(* IEC 61131-3 sources: plc-st-coding-agent/progress/evidence/f14_v14_remaining_20261113/jobs/codex_minimax-m27 (part 3) *)

(* ---- public-hard-05.patch_base_03.st ---- *)
(* ENGINEERING_CONTRACT *)
(*
  PUB001: Manual mode - button activates output while held, stop at limit switch or release.
          Manual outputs: retention=hold_until_button_release OR limit, reset=button_release OR limit_reached.
  PUB002: Emergency stop - all outputs OFF, all state cleared. No retention. Reset=EmergencyStop=TRUE.
  PUB003-PUB012: Single step mode - 8-step sequence, Start to advance each step.
          Step outputs: retention=hold_until_limit, reset=limit_reached OR mode_exit.
          Step index 1..8 maps to: Down→Grip→Up→Right→Down→Release→Up→Left→(repeat).
  PUB013-PUB014: Single cycle mode - auto-execute 8 steps on Start, stop at home.
          Same output retention as PUB003-PUB012. Cycle reset=mode_exit only.
  PUB015-PUB016: Continuous mode - same as single cycle but repeat after home.
          Cycle restart trigger: timer PT after home, if Start still asserted.
  PUB017: GripLimitSwitch/ReleaseLimitSwitch signal action completion (not position).
          Grip/Release output: activation=entry_unless_limit, retention=limit FALSE,
          deactivation=limit TRUE (same scan). No explicit reset input.
  PUB018: Caller guarantees mutually exclusive mode inputs.
  PUB019: Opposite-direction pairs (Up/Down, Left/Right) must never energize together.
          Implementation: output TRUE only when opposite limit is FALSE.
  PUB020: Single step confirmation = Start button release, not level.
*)
(* CONTRACT_RULES [] *)

TYPE ArmStep : INT (Idle := 0, Step1 := 1, Step2 := 2, Step3 := 3, Step4 := 4,
                     Step5 := 5, Step6 := 6, Step7 := 7, Step8 := 8)
END_TYPE;

FUNCTION_BLOCK ArmController
VAR_INPUT
    ManualMode       : BOOL;
    SingleStepMode   : BOOL;
    SingleCycleMode  : BOOL;
    ContinuousMode   : BOOL;
    EmergencyStop    : BOOL;
    Start            : BOOL;
    DownButton       : BOOL;
    UpButton         : BOOL;
    LeftButton       : BOOL;
    RightButton      : BOOL;
    GripButton       : BOOL;
    ReleaseButton    : BOOL;
    DownLimitSwitch  : BOOL;
    UpLimitSwitch    : BOOL;
    LeftLimitSwitch  : BOOL;
    RightLimitSwitch : BOOL;
    GripLimitSwitch  : BOOL;
    ReleaseLimitSwitch : BOOL;
END_VAR
VAR_OUTPUT
    MoveDown       : BOOL;
    MoveUp         : BOOL;
    MoveLeft       : BOOL;
    MoveRight      : BOOL;
    ActivateGrip   : BOOL;
    ActivateRelease : BOOL;
END_VAR
VAR
    tmp_CurrentStep   : ArmStep := ArmStep.Idle;
    tmp_StartTrigger  : BOOL;
    tmp_StartReleased : BOOL;
    tmp_Gripping      : BOOL;
    tmp_Releasing     : BOOL;
    tmp_CycleDoneTimer : TON;
END_VAR

// Emergency stop: clears all outputs and state
IF EmergencyStop THEN
    MoveDown       := FALSE;
    MoveUp         := FALSE;
    MoveLeft       := FALSE;
    MoveRight      := FALSE;
    ActivateGrip   := FALSE;
    ActivateRelease := FALSE;
    tmp_CurrentStep   := ArmStep.Idle;
    tmp_StartTrigger  := FALSE;
    tmp_StartReleased := FALSE;
    tmp_Gripping      := FALSE;
    tmp_Releasing     := FALSE;
    tmp_CycleDoneTimer(IN := FALSE, PT := T#0s);
    RETURN;
END_IF;

// Default all outputs OFF
MoveDown       := FALSE;
MoveUp         := FALSE;
MoveLeft       := FALSE;
MoveRight      := FALSE;
ActivateGrip   := FALSE;
ActivateRelease := FALSE;

IF ManualMode THEN
    // Direct button-to-output mapping, stop at limit switch
    MoveDown       := DownButton AND NOT DownLimitSwitch;
    MoveUp         := UpButton AND NOT UpLimitSwitch;
    MoveLeft       := LeftButton AND NOT LeftLimitSwitch;
    MoveRight      := RightButton AND NOT RightLimitSwitch;
    ActivateGrip   := GripButton AND NOT GripLimitSwitch;
    ActivateRelease := ReleaseButton AND NOT ReleaseLimitSwitch;

ELSIF SingleStepMode THEN
    // Rising-edge Start advances through steps; each step waits for limit switch
    IF tmp_StartReleased AND NOT Start AND tmp_CurrentStep = ArmStep.Idle THEN
        tmp_StartTrigger := TRUE;
    END_IF;
    tmp_StartReleased := Start;

    IF tmp_CurrentStep = ArmStep.Idle THEN
        IF tmp_StartTrigger THEN
            tmp_CurrentStep := ArmStep.Step1;
            tmp_StartTrigger := FALSE;
        END_IF;
    ELSE
        CASE TO_INT(tmp_CurrentStep) OF
            1: MoveDown := NOT DownLimitSwitch;
               IF DownLimitSwitch THEN
                   tmp_CurrentStep := ArmStep.Step2;
               END_IF;
            2: ActivateGrip := NOT GripLimitSwitch;
               IF GripLimitSwitch THEN
                   tmp_CurrentStep := ArmStep.Step3;
               END_IF;
            3: MoveUp := NOT UpLimitSwitch;
               IF UpLimitSwitch THEN
                   tmp_CurrentStep := ArmStep.Step4;
               END_IF;
            4: MoveRight := NOT RightLimitSwitch;
               IF RightLimitSwitch THEN
                   tmp_CurrentStep := ArmStep.Step5;
               END_IF;
            5: MoveDown := NOT DownLimitSwitch;
               IF DownLimitSwitch THEN
                   tmp_CurrentStep := ArmStep.Step6;
               END_IF;
            6: ActivateRelease := NOT ReleaseLimitSwitch;
               IF ReleaseLimitSwitch THEN
                   tmp_CurrentStep := ArmStep.Step7;
               END_IF;
            7: MoveUp := NOT UpLimitSwitch;
               IF UpLimitSwitch THEN
                   tmp_CurrentStep := ArmStep.Step8;
               END_IF;
            8: MoveLeft := NOT LeftLimitSwitch;
               IF LeftLimitSwitch THEN
                   tmp_CurrentStep := ArmStep.Idle;
               END_IF;
        END_CASE;
    END_IF;

ELSIF SingleCycleMode THEN
    // Start triggers auto-sequence; cycle completes and stops at home
    IF Start AND tmp_CurrentStep = ArmStep.Idle AND NOT tmp_Gripping AND NOT tmp_Releasing THEN
        tmp_StartTrigger := TRUE;
    END_IF;

    // Cycle completion: at Step8 and home (UpLimitSwitch AND LeftLimitSwitch)
    IF tmp_CurrentStep = ArmStep.Step8 AND UpLimitSwitch AND LeftLimitSwitch THEN
        tmp_CycleDoneTimer(IN := TRUE, PT := T#1ms);
        IF tmp_CycleDoneTimer.Q THEN
            tmp_StartTrigger  := FALSE;
            tmp_Gripping      := FALSE;
            tmp_Releasing     := FALSE;
            tmp_CurrentStep   := ArmStep.Idle;
        END_IF;
    ELSE
        tmp_CycleDoneTimer(IN := FALSE, PT := T#0s);
    END_IF;

    IF tmp_StartTrigger THEN
        CASE TO_INT(tmp_CurrentStep) OF
            0: tmp_CurrentStep := ArmStep.Step1;
            1: MoveDown := NOT DownLimitSwitch;
               IF DownLimitSwitch THEN
                   tmp_CurrentStep := ArmStep.Step2;
               END_IF;
            2: ActivateGrip := NOT GripLimitSwitch;
               IF GripLimitSwitch THEN
                   tmp_CurrentStep := ArmStep.Step3;
               END_IF;
            3: MoveUp := NOT UpLimitSwitch;
               IF UpLimitSwitch THEN
                   tmp_CurrentStep := ArmStep.Step4;
               END_IF;
            4: MoveRight := NOT RightLimitSwitch;
               IF RightLimitSwitch THEN
                   tmp_CurrentStep := ArmStep.Step5;
               END_IF;
            5: MoveDown := NOT DownLimitSwitch;
               IF DownLimitSwitch THEN
                   tmp_CurrentStep := ArmStep.Step6;
               END_IF;
            6: ActivateRelease := NOT ReleaseLimitSwitch;
               IF ReleaseLimitSwitch THEN
                   tmp_CurrentStep := ArmStep.Step7;
               END_IF;
            7: MoveUp := NOT UpLimitSwitch;
               IF UpLimitSwitch THEN
                   tmp_CurrentStep := ArmStep.Step8;
               END_IF;
            8: MoveLeft := NOT LeftLimitSwitch;
               IF LeftLimitSwitch THEN
                   tmp_CurrentStep := ArmStep.Idle;
               END_IF;
        END_CASE;
    END_IF;

ELSIF ContinuousMode THEN
    // Same as single cycle but restarts automatically after PT delay at home
    IF Start AND NOT tmp_Gripping AND NOT tmp_Releasing THEN
        tmp_StartTrigger := TRUE;
    END_IF;

    IF tmp_CurrentStep = ArmStep.Step8 AND UpLimitSwitch AND LeftLimitSwitch THEN
        tmp_CycleDoneTimer(IN := tmp_CycleDoneTimer.Q, PT := T#1ms);
        IF tmp_CycleDoneTimer.Q THEN
            tmp_CurrentStep := ArmStep.Idle;
        END_IF;
        IF NOT tmp_CycleDoneTimer.Q AND tmp_CurrentStep = ArmStep.Idle THEN
            tmp_StartTrigger := Start;
            tmp_Gripping     := FALSE;
            tmp_Releasing    := FALSE;
        END_IF;
    ELSE
        tmp_CycleDoneTimer(IN := FALSE, PT := T#0s);
    END_IF;

    IF tmp_StartTrigger THEN
        CASE TO_INT(tmp_CurrentStep) OF
            0: tmp_CurrentStep := ArmStep.Step1;
            1: MoveDown := NOT DownLimitSwitch;
               IF DownLimitSwitch THEN
                   tmp_CurrentStep := ArmStep.Step2;
               END_IF;
            2: ActivateGrip := NOT GripLimitSwitch;
               IF GripLimitSwitch THEN
                   tmp_CurrentStep := ArmStep.Step3;
               END_IF;
            3: MoveUp := NOT UpLimitSwitch;
               IF UpLimitSwitch THEN
                   tmp_CurrentStep := ArmStep.Step4;
               END_IF;
            4: MoveRight := NOT RightLimitSwitch;
               IF RightLimitSwitch THEN
                   tmp_CurrentStep := ArmStep.Step5;
               END_IF;
            5: MoveDown := NOT DownLimitSwitch;
               IF DownLimitSwitch THEN
                   tmp_CurrentStep := ArmStep.Step6;
               END_IF;
            6: ActivateRelease := NOT ReleaseLimitSwitch;
               IF ReleaseLimitSwitch THEN
                   tmp_CurrentStep := ArmStep.Step7;
               END_IF;
            7: MoveUp := NOT UpLimitSwitch;
               IF UpLimitSwitch THEN
                   tmp_CurrentStep := ArmStep.Step8;
               END_IF;
            8: MoveLeft := NOT LeftLimitSwitch;
               IF LeftLimitSwitch THEN
                   tmp_CurrentStep := ArmStep.Idle;
               END_IF;
        END_CASE;
    END_IF;
END_IF;

END_FUNCTION_BLOCK

(* ---- public-hard-05.raw_candidate_01.st ---- *)
(* ENGINEERING_CONTRACT *)
(*
  PUB001: Manual mode - button activates output while held, stop at limit switch or release.
          Manual outputs: retention=hold_until_button_release OR limit, reset=button_release OR limit_reached.
  PUB002: Emergency stop - all outputs OFF, all state cleared. No retention. Reset=EmergencyStop=TRUE.
  PUB003-PUB012: Single step mode - 8-step sequence, Start to advance each step.
          Step outputs: retention=hold_until_limit, reset=limit_reached OR mode_exit.
          Step index 1..8 maps to: Down→Grip→Up→Right→Down→Release→Up→Left→(repeat).
  PUB013-PUB014: Single cycle mode - auto-execute 8 steps on Start, stop at home.
          Same output retention as PUB003-PUB012. Cycle reset=mode_exit only.
  PUB015-PUB016: Continuous mode - same as single cycle but repeat after home.
          Cycle restart trigger: timer PT after home, if Start still asserted.
  PUB017: GripLimitSwitch/ReleaseLimitSwitch signal action completion (not position).
          Grip/Release output: activation=entry_unless_limit, retention=limit FALSE,
          deactivation=limit TRUE (same scan). No explicit reset input.
  PUB018: Caller guarantees mutually exclusive mode inputs.
  PUB019: Opposite-direction pairs (Up/Down, Left/Right) must never energize together.
          Implementation: output TRUE only when opposite limit is FALSE.
  PUB020: Single step confirmation = Start button release, not level.
*)
(* CONTRACT_RULES [] *)

TYPE ArmStep : INT (Idle := 0, Step1 := 1, Step2 := 2, Step3 := 3, Step4 := 4,
                     Step5 := 5, Step6 := 6, Step7 := 7, Step8 := 8)
END_TYPE

FUNCTION_BLOCK ArmController
VAR_INPUT
    ManualMode       : BOOL;
    SingleStepMode   : BOOL;
    SingleCycleMode  : BOOL;
    ContinuousMode   : BOOL;
    EmergencyStop    : BOOL;
    Start            : BOOL;
    DownButton       : BOOL;
    UpButton         : BOOL;
    LeftButton       : BOOL;
    RightButton      : BOOL;
    GripButton       : BOOL;
    ReleaseButton    : BOOL;
    DownLimitSwitch  : BOOL;
    UpLimitSwitch    : BOOL;
    LeftLimitSwitch  : BOOL;
    RightLimitSwitch : BOOL;
    GripLimitSwitch  : BOOL;
    ReleaseLimitSwitch : BOOL;
END_VAR
VAR_OUTPUT
    MoveDown       : BOOL;
    MoveUp         : BOOL;
    MoveLeft       : BOOL;
    MoveRight      : BOOL;
    ActivateGrip   : BOOL;
    ActivateRelease : BOOL;
END_VAR
VAR
    tmp_CurrentStep   : ArmStep := ArmStep.Idle;
    tmp_StartTrigger  : BOOL;
    tmp_StartReleased : BOOL;
    tmp_Gripping      : BOOL;
    tmp_Releasing     : BOOL;
    tmp_CycleDoneTimer : TON;
END_VAR

// Emergency stop: clears all outputs and state
IF EmergencyStop THEN
    MoveDown       := FALSE;
    MoveUp         := FALSE;
    MoveLeft       := FALSE;
    MoveRight      := FALSE;
    ActivateGrip   := FALSE;
    ActivateRelease := FALSE;
    tmp_CurrentStep   := ArmStep.Idle;
    tmp_StartTrigger  := FALSE;
    tmp_StartReleased := FALSE;
    tmp_Gripping      := FALSE;
    tmp_Releasing     := FALSE;
    tmp_CycleDoneTimer(IN := FALSE, PT := T#0s);
    RETURN;
END_IF;

// Default all outputs OFF
MoveDown       := FALSE;
MoveUp         := FALSE;
MoveLeft       := FALSE;
MoveRight      := FALSE;
ActivateGrip   := FALSE;
ActivateRelease := FALSE;

IF ManualMode THEN
    // Direct button-to-output mapping, stop at limit switch
    MoveDown       := DownButton AND NOT DownLimitSwitch;
    MoveUp         := UpButton AND NOT UpLimitSwitch;
    MoveLeft       := LeftButton AND NOT LeftLimitSwitch;
    MoveRight      := RightButton AND NOT RightLimitSwitch;
    ActivateGrip   := GripButton AND NOT GripLimitSwitch;
    ActivateRelease := ReleaseButton AND NOT ReleaseLimitSwitch;

ELSIF SingleStepMode THEN
    // Rising-edge Start advances through steps; each step waits for limit switch
    IF tmp_StartReleased AND NOT Start AND tmp_CurrentStep = ArmStep.Idle THEN
        tmp_StartTrigger := TRUE;
    END_IF
    tmp_StartReleased := Start;

    IF tmp_CurrentStep = ArmStep.Idle THEN
        IF tmp_StartTrigger THEN
            tmp_CurrentStep := ArmStep.Step1;
            tmp_StartTrigger := FALSE;
        END_IF;
    ELSE
        CASE TO_INT(tmp_CurrentStep) OF
            1: MoveDown := NOT DownLimitSwitch;
               IF DownLimitSwitch THEN
                   tmp_CurrentStep := ArmStep.Step2;
               END_IF;
            2: ActivateGrip := NOT GripLimitSwitch;
               IF GripLimitSwitch THEN
                   tmp_CurrentStep := ArmStep.Step3;
               END_IF;
            3: MoveUp := NOT UpLimitSwitch;
               IF UpLimitSwitch THEN
                   tmp_CurrentStep := ArmStep.Step4;
               END_IF;
            4: MoveRight := NOT RightLimitSwitch;
               IF RightLimitSwitch THEN
                   tmp_CurrentStep := ArmStep.Step5;
               END_IF;
            5: MoveDown := NOT DownLimitSwitch;
               IF DownLimitSwitch THEN
                   tmp_CurrentStep := ArmStep.Step6;
               END_IF;
            6: ActivateRelease := NOT ReleaseLimitSwitch;
               IF ReleaseLimitSwitch THEN
                   tmp_CurrentStep := ArmStep.Step7;
               END_IF;
            7: MoveUp := NOT UpLimitSwitch;
               IF UpLimitSwitch THEN
                   tmp_CurrentStep := ArmStep.Step8;
               END_IF;
            8: MoveLeft := NOT LeftLimitSwitch;
               IF LeftLimitSwitch THEN
                   tmp_CurrentStep := ArmStep.Idle;
               END_IF;
        END_CASE;
    END_IF;

ELSIF SingleCycleMode THEN
    // Start triggers auto-sequence; cycle completes and stops at home
    IF Start AND tmp_CurrentStep = ArmStep.Idle AND NOT tmp_Gripping AND NOT tmp_Releasing THEN
        tmp_StartTrigger := TRUE;
    END_IF;

    // Cycle completion: at Step8 and home (UpLimitSwitch AND LeftLimitSwitch)
    IF tmp_CurrentStep = ArmStep.Step8 AND UpLimitSwitch AND LeftLimitSwitch THEN
        tmp_CycleDoneTimer(IN := TRUE, PT := T#1ms);
        IF tmp_CycleDoneTimer.Q THEN
            tmp_StartTrigger  := FALSE;
            tmp_Gripping      := FALSE;
            tmp_Releasing     := FALSE;
            tmp_CurrentStep   := ArmStep.Idle;
        END_IF;
    ELSE
        tmp_CycleDoneTimer(IN := FALSE, PT := T#0s);
    END_IF;

    IF tmp_StartTrigger THEN
        CASE TO_INT(tmp_CurrentStep) OF
            0: tmp_CurrentStep := ArmStep.Step1;
            1: MoveDown := NOT DownLimitSwitch;
               IF DownLimitSwitch THEN
                   tmp_CurrentStep := ArmStep.Step2;
               END_IF;
            2: ActivateGrip := NOT GripLimitSwitch;
               IF GripLimitSwitch THEN
                   tmp_CurrentStep := ArmStep.Step3;
               END_IF;
            3: MoveUp := NOT UpLimitSwitch;
               IF UpLimitSwitch THEN
                   tmp_CurrentStep := ArmStep.Step4;
               END_IF;
            4: MoveRight := NOT RightLimitSwitch;
               IF RightLimitSwitch THEN
                   tmp_CurrentStep := ArmStep.Step5;
               END_IF;
            5: MoveDown := NOT DownLimitSwitch;
               IF DownLimitSwitch THEN
                   tmp_CurrentStep := ArmStep.Step6;
               END_IF;
            6: ActivateRelease := NOT ReleaseLimitSwitch;
               IF ReleaseLimitSwitch THEN
                   tmp_CurrentStep := ArmStep.Step7;
               END_IF;
            7: MoveUp := NOT UpLimitSwitch;
               IF UpLimitSwitch THEN
                   tmp_CurrentStep := ArmStep.Step8;
               END_IF;
            8: MoveLeft := NOT LeftLimitSwitch;
               IF LeftLimitSwitch THEN
                   tmp_CurrentStep := ArmStep.Idle;
               END_IF;
        END_CASE;
    END_IF;

ELSIF ContinuousMode THEN
    // Same as single cycle but restarts automatically after PT delay at home
    IF Start AND NOT tmp_Gripping AND NOT tmp_Releasing THEN
        tmp_StartTrigger := TRUE;
    END_IF;

    IF tmp_CurrentStep = ArmStep.Step8 AND UpLimitSwitch AND LeftLimitSwitch THEN
        tmp_CycleDoneTimer(IN := tmp_CycleDoneTimer.Q, PT := T#1ms);
        IF tmp_CycleDoneTimer.Q THEN
            tmp_CurrentStep := ArmStep.Idle;
        END_IF;
        IF NOT tmp_CycleDoneTimer.Q AND tmp_CurrentStep = ArmStep.Idle THEN
            tmp_StartTrigger := Start;
            tmp_Gripping     := FALSE;
            tmp_Releasing    := FALSE;
        END_IF;
    ELSE
        tmp_CycleDoneTimer(IN := FALSE, PT := T#0s);
    END_IF;

    IF tmp_StartTrigger THEN
        CASE TO_INT(tmp_CurrentStep) OF
            0: tmp_CurrentStep := ArmStep.Step1;
            1: MoveDown := NOT DownLimitSwitch;
               IF DownLimitSwitch THEN
                   tmp_CurrentStep := ArmStep.Step2;
               END_IF;
            2: ActivateGrip := NOT GripLimitSwitch;
               IF GripLimitSwitch THEN
                   tmp_CurrentStep := ArmStep.Step3;
               END_IF;
            3: MoveUp := NOT UpLimitSwitch;
               IF UpLimitSwitch THEN
                   tmp_CurrentStep := ArmStep.Step4;
               END_IF;
            4: MoveRight := NOT RightLimitSwitch;
               IF RightLimitSwitch THEN
                   tmp_CurrentStep := ArmStep.Step5;
               END_IF;
            5: MoveDown := NOT DownLimitSwitch;
               IF DownLimitSwitch THEN
                   tmp_CurrentStep := ArmStep.Step6;
               END_IF;
            6: ActivateRelease := NOT ReleaseLimitSwitch;
               IF ReleaseLimitSwitch THEN
                   tmp_CurrentStep := ArmStep.Step7;
               END_IF;
            7: MoveUp := NOT UpLimitSwitch;
               IF UpLimitSwitch THEN
                   tmp_CurrentStep := ArmStep.Step8;
               END_IF;
            8: MoveLeft := NOT LeftLimitSwitch;
               IF LeftLimitSwitch THEN
                   tmp_CurrentStep := ArmStep.Idle;
               END_IF;
        END_CASE;
    END_IF;
END_IF;

END_FUNCTION_BLOCK

(* ---- public-hard-06.candidate_01.st ---- *)
(*
ENGINEERING_CONTRACT
===================
PUB001: Mode 0=Manual, 1=Automatic (VAR_INPUT Mode)
PUB003: Manual interlock - ForwardButton→MotorForward, ReverseButton→MotorReverse, mutually exclusive
PUB002: Automatic sequential transport: Feed→Wash→Weigh→Fire→Output stations
PUB004: Station arrival detected by sensors; motor stops, awaits completion signal, then advances
PUB006: Weight qualification: qualified if 100<=weight<=200; else kick initiated
PUB007: FiringTemp calculation: weight[100,200]→temp[500,550] via linear interpolation
PUB008: CompletionLight ON when product detected at output, OFF when product removed
PUB005/P UB009-PUB012: washComplete/weightComplete/firingComplete are external process signals

OUTPUT STATE RETENTION
- MotorForward/MotorReverse: combinational per Mode selection, no retention across modes
- kick: pulse on weight qualification failure, no hold required
- CompletionLight: retained based on SensorOutput (hold until product removed)
- firingTemp: retained value written at weight station, held through firing until output

SCAN BEHAVIOR
- Sequential automatic states evaluate same-scan final state before output
- TON not required; all timing handled externally via completion signals
- Direction rule: MotorForward and MotorReverse never energized together
*)

FUNCTION_BLOCK ProductionControl
VAR_INPUT
    Mode            : BOOL;
    ForwardButton   : BOOL;
    ReverseButton   : BOOL;
    SensorFeed      : BOOL;
    SensorWash      : BOOL;
    SensorWeight    : BOOL;
    SensorFiring    : BOOL;
    SensorOutput    : BOOL;
    washComplete    : BOOL;
    weightComplete  : BOOL;
    weight          : REAL;
    firingComplete  : BOOL;
END_VAR

VAR_OUTPUT
    MotorForward    : BOOL;
    MotorReverse    : BOOL;
    kick             : BOOL;
    CompletionLight  : BOOL;
    firingTemp       : REAL;
END_VAR

VAR
    stepPosition    : INT := 0;
    localKick       : BOOL := FALSE;
END_VAR

(* CONTRACT_RULES [] *)

CASE stepPosition OF
    0: (* At feed station - waiting for material *)
        IF SensorFeed THEN
            MotorForward := TRUE;
            stepPosition := 1;
        END_IF;

    1: (* Moving to wash station - detecting arrival *)
        IF SensorWash THEN
            MotorForward := FALSE;
            stepPosition := 2;
        END_IF;

    2: (* At wash station - waiting for washComplete *)
        IF washComplete THEN
            MotorForward := TRUE;
            stepPosition := 3;
        END_IF;

    3: (* Moving to weight station - detecting arrival *)
        IF SensorWeight THEN
            MotorForward := FALSE;
            stepPosition := 4;
        END_IF;

    4: (* At weight station - waiting for weightComplete *)
        IF weightComplete THEN
            IF (weight >= 100.0) AND (weight <= 200.0) THEN
                firingTemp := 500.0 + (weight - 100.0) * (50.0 / 100.0);
                MotorForward := TRUE;
                stepPosition := 5;
            ELSE
                localKick := TRUE;
                kick := TRUE;
                MotorReverse := TRUE;
                stepPosition := 6;
            END_IF;
        END_IF;

    5: (* Moving to firing station - detecting arrival *)
        IF SensorFiring THEN
            MotorForward := FALSE;
            stepPosition := 7;
        END_IF;

    6: (* Rejection - returning to feed station *)
        localKick := FALSE;
        kick := FALSE;
        IF NOT SensorFeed THEN
            MotorReverse := FALSE;
            stepPosition := 0;
        END_IF;

    7: (* At firing station - waiting for firingComplete *)
        IF firingComplete THEN
            MotorForward := TRUE;
            stepPosition := 8;
        END_IF;

    8: (* Moving to output station - detecting arrival *)
        IF SensorOutput THEN
            MotorForward := FALSE;
            stepPosition := 9;
        END_IF;

    9: (* At output station - waiting for product removal *)
        CompletionLight := TRUE;

    ELSE
        stepPosition := 0;
END_CASE;

IF Mode = 0 THEN
    stepPosition := 0;
    MotorForward := FALSE;
    MotorReverse := FALSE;
    kick := FALSE;
    CompletionLight := FALSE;
    localKick := FALSE;
    firingTemp := 0.0;

    IF ForwardButton AND NOT ReverseButton THEN
        MotorForward := TRUE;
    ELSIF ReverseButton AND NOT ForwardButton THEN
        MotorReverse := TRUE;
    END_IF;
END_IF;

IF NOT SensorOutput AND stepPosition = 9 THEN
    CompletionLight := FALSE;
    stepPosition := 0;
END_IF;

END_FUNCTION_BLOCK

(* ---- public-hard-06.raw_candidate_01.st ---- *)
(*
ENGINEERING_CONTRACT
===================
PUB001: Mode 0=Manual, 1=Automatic (VAR_INPUT Mode)
PUB003: Manual interlock - ForwardButton→MotorForward, ReverseButton→MotorReverse, mutually exclusive
PUB002: Automatic sequential transport: Feed→Wash→Weigh→Fire→Output stations
PUB004: Station arrival detected by sensors; motor stops, awaits completion signal, then advances
PUB006: Weight qualification: qualified if 100<=weight<=200; else kick initiated
PUB007: FiringTemp calculation: weight[100,200]→temp[500,550] via linear interpolation
PUB008: CompletionLight ON when product detected at output, OFF when product removed
PUB005/P UB009-PUB012: washComplete/weightComplete/firingComplete are external process signals

OUTPUT STATE RETENTION
- MotorForward/MotorReverse: combinational per Mode selection, no retention across modes
- kick: pulse on weight qualification failure, no hold required
- CompletionLight: retained based on SensorOutput (hold until product removed)
- firingTemp: retained value written at weight station, held through firing until output

SCAN BEHAVIOR
- Sequential automatic states evaluate same-scan final state before output
- TON not required; all timing handled externally via completion signals
- Direction rule: MotorForward and MotorReverse never energized together
*)

FUNCTION_BLOCK ProductionControl
VAR_INPUT
    Mode            : BOOL;
    ForwardButton   : BOOL;
    ReverseButton   : BOOL;
    SensorFeed      : BOOL;
    SensorWash      : BOOL;
    SensorWeight    : BOOL;
    SensorFiring    : BOOL;
    SensorOutput    : BOOL;
    washComplete    : BOOL;
    weightComplete  : BOOL;
    weight          : REAL;
    firingComplete  : BOOL;
END_VAR

VAR_OUTPUT
    MotorForward    : BOOL;
    MotorReverse    : BOOL;
    kick             : BOOL;
    CompletionLight  : BOOL;
    firingTemp       : REAL;
END_VAR

VAR
    stepPosition    : INT := 0;
    localKick       : BOOL := FALSE;
END_VAR

(* CONTRACT_RULES [] *)

CASE stepPosition OF
    0: (* At feed station - waiting for material *)
        IF SensorFeed THEN
            MotorForward := TRUE;
            stepPosition := 1;
        END_IF

    1: (* Moving to wash station - detecting arrival *)
        IF SensorWash THEN
            MotorForward := FALSE;
            stepPosition := 2;
        END_IF

    2: (* At wash station - waiting for washComplete *)
        IF washComplete THEN
            MotorForward := TRUE;
            stepPosition := 3;
        END_IF

    3: (* Moving to weight station - detecting arrival *)
        IF SensorWeight THEN
            MotorForward := FALSE;
            stepPosition := 4;
        END_IF

    4: (* At weight station - waiting for weightComplete *)
        IF weightComplete THEN
            IF (weight >= 100.0) AND (weight <= 200.0) THEN
                firingTemp := 500.0 + (weight - 100.0) * (50.0 / 100.0);
                MotorForward := TRUE;
                stepPosition := 5;
            ELSE
                localKick := TRUE;
                kick := TRUE;
                MotorReverse := TRUE;
                stepPosition := 6;
            END_IF
        END_IF

    5: (* Moving to firing station - detecting arrival *)
        IF SensorFiring THEN
            MotorForward := FALSE;
            stepPosition := 7;
        END_IF

    6: (* Rejection - returning to feed station *)
        localKick := FALSE;
        kick := FALSE;
        IF NOT SensorFeed THEN
            MotorReverse := FALSE;
            stepPosition := 0;
        END_IF

    7: (* At firing station - waiting for firingComplete *)
        IF firingComplete THEN
            MotorForward := TRUE;
            stepPosition := 8;
        END_IF

    8: (* Moving to output station - detecting arrival *)
        IF SensorOutput THEN
            MotorForward := FALSE;
            stepPosition := 9;
        END_IF

    9: (* At output station - waiting for product removal *)
        CompletionLight := TRUE;

    ELSE
        stepPosition := 0;
END_CASE

IF Mode = 0 THEN
    stepPosition := 0;
    MotorForward := FALSE;
    MotorReverse := FALSE;
    kick := FALSE;
    CompletionLight := FALSE;
    localKick := FALSE;
    firingTemp := 0.0;

    IF ForwardButton AND NOT ReverseButton THEN
        MotorForward := TRUE;
    ELSIF ReverseButton AND NOT ForwardButton THEN
        MotorReverse := TRUE;
    END_IF
END_IF

IF NOT SensorOutput AND stepPosition = 9 THEN
    CompletionLight := FALSE;
    stepPosition := 0;
END_IF

END_FUNCTION_BLOCK

(* ---- public-medium-01.candidate_01.st ---- *)
FUNCTION_BLOCK FB_MultiPumpControl
VAR_INPUT
    mode : BOOL;          // FALSE: Manual mode, TRUE: Automatic mode
    start : BOOL;         // Start button
    stop : BOOL;          // Stop button
END_VAR

VAR_IN_OUT
    pumpGroup : ARRAY[1..5] OF ST_Pump;
END_VAR

VAR
    startRisingEdge : BOOL;               // Rising edge of start
    tmp_startPrev : BOOL;                 // Previous start state
    tmp_i : INT;                          // Loop counter
    tmp_j : INT;                          // Loop counter
    tmp_swap : INT;                       // Swap variable
    tmp_pumpIdx : ARRAY[1..5] OF INT;    // Pump indices for sorting
    tmp_priorities : ARRAY[1..5] OF INT; // Priority copy for sorting
    tmp_swap_idx : INT;                   // Index swap
END_VAR

// ENGINEERING_CONTRACT:
// PUB001 [L91-265]: mode=FALSE → manual; start activates pumps where selection=TRUE
// PUB001 [L91-265]: mode=TRUE → automatic; start activates top-3 by priority (3-in-2-standby)
// PUB002 [L266-350]: stop halts all pumps; no retention on stop (level-triggered)
// PUB003 [L351-463]: Rising edge on start evaluates selection; stop has same-scan priority
// PUB004 [L464-652]: Only RunComd is written; priority/selection are read-only

(* CONTRACT_RULES [] *)

startRisingEdge := start AND NOT tmp_startPrev;

IF stop THEN
    FOR tmp_i := 1 TO 5 DO
        pumpGroup[tmp_i].RunComd := FALSE;
    END_FOR;
ELSIF startRisingEdge THEN
    IF mode = FALSE THEN
        FOR tmp_i := 1 TO 5 DO
            IF pumpGroup[tmp_i].selection THEN
                pumpGroup[tmp_i].RunComd := TRUE;
            END_IF;
        END_FOR;
    ELSE
        FOR tmp_i := 1 TO 5 DO
            tmp_priorities[tmp_i] := pumpGroup[tmp_i].priority;
            tmp_pumpIdx[tmp_i] := tmp_i;
        END_FOR;
        FOR tmp_i := 1 TO 4 DO
            FOR tmp_j := tmp_i + 1 TO 5 DO
                IF tmp_priorities[tmp_j] > tmp_priorities[tmp_i] THEN
                    tmp_swap := tmp_priorities[tmp_i];
                    tmp_priorities[tmp_i] := tmp_priorities[tmp_j];
                    tmp_priorities[tmp_j] := tmp_swap;
                    tmp_swap_idx := tmp_pumpIdx[tmp_i];
                    tmp_pumpIdx[tmp_i] := tmp_pumpIdx[tmp_j];
                    tmp_pumpIdx[tmp_j] := tmp_swap_idx;
                END_IF;
            END_FOR;
        END_FOR;
        FOR tmp_i := 1 TO 5 DO
            IF tmp_i <= 3 THEN
                pumpGroup[tmp_pumpIdx[tmp_i]].RunComd := TRUE;
            ELSE
                pumpGroup[tmp_pumpIdx[tmp_i]].RunComd := FALSE;
            END_IF;
        END_FOR;
    END_IF;
END_IF;

tmp_startPrev := start;
END_FUNCTION_BLOCK

(* ---- public-medium-01.candidate_03.st ---- *)
TYPE ST_Pump :
STRUCT
    priority : INT;
    selection : BOOL;
    RunComd : BOOL;
END_STRUCT
END_TYPE;

FUNCTION_BLOCK FB_MultiPumpControl
VAR_INPUT
    mode : BOOL;          // FALSE: Manual mode, TRUE: Automatic mode
    start : BOOL;         // Start button
    stop : BOOL;          // Stop button
END_VAR

VAR_IN_OUT
    pumpGroup : ARRAY[1..5] OF ST_Pump;
END_VAR

VAR
    startRisingEdge : BOOL;               // Rising edge of start
    tmp_startPrev : BOOL;                 // Previous start state
    tmp_i : INT;                          // Loop counter
    tmp_j : INT;                          // Loop counter
    tmp_swap : INT;                       // Swap variable
    tmp_pumpIdx : ARRAY[1..5] OF INT;    // Pump indices for sorting
    tmp_priorities : ARRAY[1..5] OF INT; // Priority copy for sorting
    tmp_swap_idx : INT;                   // Index swap
END_VAR

// ENGINEERING_CONTRACT:
// PUB001 [L91-265]: mode=FALSE → manual; start activates pumps where selection=TRUE
// PUB001 [L91-265]: mode=TRUE → automatic; start activates top-3 by priority (3-in-2-standby)
// PUB002 [L266-350]: stop halts all pumps; no retention on stop (level-triggered)
// PUB003 [L351-463]: Rising edge on start evaluates selection; stop has same-scan priority
// PUB004 [L464-652]: Only RunComd is written; priority/selection are read-only

(* CONTRACT_RULES [] *)

startRisingEdge := start AND NOT tmp_startPrev;

IF stop THEN
    FOR tmp_i := 1 TO 5 DO
        pumpGroup[tmp_i].RunComd := FALSE;
    END_FOR;
ELSIF startRisingEdge THEN
    IF mode = FALSE THEN
        FOR tmp_i := 1 TO 5 DO
            IF pumpGroup[tmp_i].selection THEN
                pumpGroup[tmp_i].RunComd := TRUE;
            END_IF;
        END_FOR;
    ELSE
        FOR tmp_i := 1 TO 5 DO
            tmp_priorities[tmp_i] := pumpGroup[tmp_i].priority;
            tmp_pumpIdx[tmp_i] := tmp_i;
        END_FOR;
        FOR tmp_i := 1 TO 4 DO
            FOR tmp_j := tmp_i + 1 TO 5 DO
                IF tmp_priorities[tmp_j] > tmp_priorities[tmp_i] THEN
                    tmp_swap := tmp_priorities[tmp_i];
                    tmp_priorities[tmp_i] := tmp_priorities[tmp_j];
                    tmp_priorities[tmp_j] := tmp_swap;
                    tmp_swap_idx := tmp_pumpIdx[tmp_i];
                    tmp_pumpIdx[tmp_i] := tmp_pumpIdx[tmp_j];
                    tmp_pumpIdx[tmp_j] := tmp_swap_idx;
                END_IF;
            END_FOR;
        END_FOR;
        FOR tmp_i := 1 TO 5 DO
            IF tmp_i <= 3 THEN
                pumpGroup[tmp_pumpIdx[tmp_i]].RunComd := TRUE;
            ELSE
                pumpGroup[tmp_pumpIdx[tmp_i]].RunComd := FALSE;
            END_IF;
        END_FOR;
    END_IF;
END_IF;

tmp_startPrev := start;
END_FUNCTION_BLOCK

(* ---- public-medium-01.patch_base_02.st ---- *)
FUNCTION_BLOCK FB_MultiPumpControl
VAR_INPUT
    mode : BOOL;          // FALSE: Manual mode, TRUE: Automatic mode
    start : BOOL;         // Start button
    stop : BOOL;          // Stop button
END_VAR

VAR_IN_OUT
    pumpGroup : ARRAY[1..5] OF ST_Pump;
END_VAR

VAR
    startRisingEdge : BOOL;               // Rising edge of start
    tmp_startPrev : BOOL;                 // Previous start state
    tmp_i : INT;                          // Loop counter
    tmp_j : INT;                          // Loop counter
    tmp_swap : INT;                       // Swap variable
    tmp_pumpIdx : ARRAY[1..5] OF INT;    // Pump indices for sorting
    tmp_priorities : ARRAY[1..5] OF INT; // Priority copy for sorting
    tmp_swap_idx : INT;                   // Index swap
END_VAR

// ENGINEERING_CONTRACT:
// PUB001 [L91-265]: mode=FALSE → manual; start activates pumps where selection=TRUE
// PUB001 [L91-265]: mode=TRUE → automatic; start activates top-3 by priority (3-in-2-standby)
// PUB002 [L266-350]: stop halts all pumps; no retention on stop (level-triggered)
// PUB003 [L351-463]: Rising edge on start evaluates selection; stop has same-scan priority
// PUB004 [L464-652]: Only RunComd is written; priority/selection are read-only

(* CONTRACT_RULES [] *)

startRisingEdge := start AND NOT tmp_startPrev;

IF stop THEN
    FOR tmp_i := 1 TO 5 DO
        pumpGroup[tmp_i].RunComd := FALSE;
    END_FOR;
ELSIF startRisingEdge THEN
    IF mode = FALSE THEN
        FOR tmp_i := 1 TO 5 DO
            IF pumpGroup[tmp_i].selection THEN
                pumpGroup[tmp_i].RunComd := TRUE;
            END_IF;
        END_FOR;
    ELSE
        FOR tmp_i := 1 TO 5 DO
            tmp_priorities[tmp_i] := pumpGroup[tmp_i].priority;
            tmp_pumpIdx[tmp_i] := tmp_i;
        END_FOR;
        FOR tmp_i := 1 TO 4 DO
            FOR tmp_j := tmp_i + 1 TO 5 DO
                IF tmp_priorities[tmp_j] > tmp_priorities[tmp_i] THEN
                    tmp_swap := tmp_priorities[tmp_i];
                    tmp_priorities[tmp_i] := tmp_priorities[tmp_j];
                    tmp_priorities[tmp_j] := tmp_swap;
                    tmp_swap_idx := tmp_pumpIdx[tmp_i];
                    tmp_pumpIdx[tmp_i] := tmp_pumpIdx[tmp_j];
                    tmp_pumpIdx[tmp_j] := tmp_swap_idx;
                END_IF;
            END_FOR;
        END_FOR;
        FOR tmp_i := 1 TO 5 DO
            IF tmp_i <= 3 THEN
                pumpGroup[tmp_pumpIdx[tmp_i]].RunComd := TRUE;
            ELSE
                pumpGroup[tmp_pumpIdx[tmp_i]].RunComd := FALSE;
            END_IF;
        END_FOR;
    END_IF;
END_IF;

tmp_startPrev := start;
END_FUNCTION_BLOCK

(* ---- public-medium-01.patch_base_03.st ---- *)
FUNCTION_BLOCK FB_MultiPumpControl
VAR_INPUT
    mode : BOOL;          // FALSE: Manual mode, TRUE: Automatic mode
    start : BOOL;         // Start button
    stop : BOOL;          // Stop button
END_VAR

VAR_IN_OUT
    pumpGroup : ARRAY[1..5] OF ST_Pump;
END_VAR

VAR
    startRisingEdge : BOOL;               // Rising edge of start
    tmp_startPrev : BOOL;                 // Previous start state
    tmp_i : INT;                          // Loop counter
    tmp_j : INT;                          // Loop counter
    tmp_swap : INT;                       // Swap variable
    tmp_pumpIdx : ARRAY[1..5] OF INT;    // Pump indices for sorting
    tmp_priorities : ARRAY[1..5] OF INT; // Priority copy for sorting
    tmp_swap_idx : INT;                   // Index swap
END_VAR

// ENGINEERING_CONTRACT:
// PUB001 [L91-265]: mode=FALSE → manual; start activates pumps where selection=TRUE
// PUB001 [L91-265]: mode=TRUE → automatic; start activates top-3 by priority (3-in-2-standby)
// PUB002 [L266-350]: stop halts all pumps; no retention on stop (level-triggered)
// PUB003 [L351-463]: Rising edge on start evaluates selection; stop has same-scan priority
// PUB004 [L464-652]: Only RunComd is written; priority/selection are read-only

(* CONTRACT_RULES [] *)

startRisingEdge := start AND NOT tmp_startPrev;

IF stop THEN
    FOR tmp_i := 1 TO 5 DO
        pumpGroup[tmp_i].RunComd := FALSE;
    END_FOR;
ELSIF startRisingEdge THEN
    IF mode = FALSE THEN
        FOR tmp_i := 1 TO 5 DO
            IF pumpGroup[tmp_i].selection THEN
                pumpGroup[tmp_i].RunComd := TRUE;
            END_IF;
        END_FOR;
    ELSE
        FOR tmp_i := 1 TO 5 DO
            tmp_priorities[tmp_i] := pumpGroup[tmp_i].priority;
            tmp_pumpIdx[tmp_i] := tmp_i;
        END_FOR;
        FOR tmp_i := 1 TO 4 DO
            FOR tmp_j := tmp_i + 1 TO 5 DO
                IF tmp_priorities[tmp_j] > tmp_priorities[tmp_i] THEN
                    tmp_swap := tmp_priorities[tmp_i];
                    tmp_priorities[tmp_i] := tmp_priorities[tmp_j];
                    tmp_priorities[tmp_j] := tmp_swap;
                    tmp_swap_idx := tmp_pumpIdx[tmp_i];
                    tmp_pumpIdx[tmp_i] := tmp_pumpIdx[tmp_j];
                    tmp_pumpIdx[tmp_j] := tmp_swap_idx;
                END_IF;
            END_FOR;
        END_FOR;
        FOR tmp_i := 1 TO 5 DO
            IF tmp_i <= 3 THEN
                pumpGroup[tmp_pumpIdx[tmp_i]].RunComd := TRUE;
            ELSE
                pumpGroup[tmp_pumpIdx[tmp_i]].RunComd := FALSE;
            END_IF;
        END_FOR;
    END_IF;
END_IF;

tmp_startPrev := start;
END_FUNCTION_BLOCK

(* ---- public-medium-01.patch_base_04.st ---- *)
TYPE ST_Pump :
STRUCT
    priority : INT;
    selection : BOOL;
    RunComd : BOOL;
END_STRUCT
END_TYPE;

FUNCTION_BLOCK FB_MultiPumpControl
VAR_INPUT
    mode : BOOL;          // FALSE: Manual mode, TRUE: Automatic mode
    start : BOOL;         // Start button
    stop : BOOL;          // Stop button
END_VAR

VAR_IN_OUT
    pumpGroup : ARRAY[1..5] OF ST_Pump;
END_VAR

VAR
    startRisingEdge : BOOL;               // Rising edge of start
    tmp_startPrev : BOOL;                 // Previous start state
    tmp_i : INT;                          // Loop counter
    tmp_j : INT;                          // Loop counter
    tmp_swap : INT;                       // Swap variable
    tmp_pumpIdx : ARRAY[1..5] OF INT;    // Pump indices for sorting
    tmp_priorities : ARRAY[1..5] OF INT; // Priority copy for sorting
    tmp_swap_idx : INT;                   // Index swap
END_VAR

// ENGINEERING_CONTRACT:
// PUB001 [L91-265]: mode=FALSE → manual; start activates pumps where selection=TRUE
// PUB001 [L91-265]: mode=TRUE → automatic; start activates top-3 by priority (3-in-2-standby)
// PUB002 [L266-350]: stop halts all pumps; no retention on stop (level-triggered)
// PUB003 [L351-463]: Rising edge on start evaluates selection; stop has same-scan priority
// PUB004 [L464-652]: Only RunComd is written; priority/selection are read-only

(* CONTRACT_RULES [] *)

startRisingEdge := start AND NOT tmp_startPrev;

IF stop THEN
    FOR tmp_i := 1 TO 5 DO
        pumpGroup[tmp_i].RunComd := FALSE;
    END_FOR;
ELSIF startRisingEdge THEN
    IF mode = FALSE THEN
        FOR tmp_i := 1 TO 5 DO
            IF pumpGroup[tmp_i].selection THEN
                pumpGroup[tmp_i].RunComd := TRUE;
            END_IF;
        END_FOR;
    ELSE
        FOR tmp_i := 1 TO 5 DO
            tmp_priorities[tmp_i] := pumpGroup[tmp_i].priority;
            tmp_pumpIdx[tmp_i] := tmp_i;
        END_FOR;
        FOR tmp_i := 1 TO 4 DO
            FOR tmp_j := tmp_i + 1 TO 5 DO
                IF tmp_priorities[tmp_j] > tmp_priorities[tmp_i] THEN
                    tmp_swap := tmp_priorities[tmp_i];
                    tmp_priorities[tmp_i] := tmp_priorities[tmp_j];
                    tmp_priorities[tmp_j] := tmp_swap;
                    tmp_swap_idx := tmp_pumpIdx[tmp_i];
                    tmp_pumpIdx[tmp_i] := tmp_pumpIdx[tmp_j];
                    tmp_pumpIdx[tmp_j] := tmp_swap_idx;
                END_IF;
            END_FOR;
        END_FOR;
        FOR tmp_i := 1 TO 5 DO
            IF tmp_i <= 3 THEN
                pumpGroup[tmp_pumpIdx[tmp_i]].RunComd := TRUE;
            ELSE
                pumpGroup[tmp_pumpIdx[tmp_i]].RunComd := FALSE;
            END_IF;
        END_FOR;
    END_IF;
END_IF;

tmp_startPrev := start;
END_FUNCTION_BLOCK

(* ---- public-medium-01.raw_candidate_01.st ---- *)
FUNCTION_BLOCK FB_MultiPumpControl
VAR_INPUT
    mode : BOOL;          // FALSE: Manual mode, TRUE: Automatic mode
    start : BOOL;         // Start button
    stop : BOOL;          // Stop button
END_VAR

VAR_IN_OUT
    pumpGroup : ARRAY[1..5] OF ST_Pump;
END_VAR

VAR
    startRisingEdge : BOOL;               // Rising edge of start
    tmp_startPrev : BOOL;                 // Previous start state
    tmp_i : INT;                          // Loop counter
    tmp_j : INT;                          // Loop counter
    tmp_swap : INT;                       // Swap variable
    tmp_pumpIdx : ARRAY[1..5] OF INT;    // Pump indices for sorting
    tmp_priorities : ARRAY[1..5] OF INT; // Priority copy for sorting
    tmp_swap_idx : INT;                   // Index swap
END_VAR

// ENGINEERING_CONTRACT:
// PUB001 [L91-265]: mode=FALSE → manual; start activates pumps where selection=TRUE
// PUB001 [L91-265]: mode=TRUE → automatic; start activates top-3 by priority (3-in-2-standby)
// PUB002 [L266-350]: stop halts all pumps; no retention on stop (level-triggered)
// PUB003 [L351-463]: Rising edge on start evaluates selection; stop has same-scan priority
// PUB004 [L464-652]: Only RunComd is written; priority/selection are read-only

(* CONTRACT_RULES [] *)

startRisingEdge := start AND NOT tmp_startPrev;

IF stop THEN
    FOR tmp_i := 1 TO 5 DO
        pumpGroup[tmp_i].RunComd := FALSE;
    END_FOR
ELSIF startRisingEdge THEN
    IF mode = FALSE THEN
        FOR tmp_i := 1 TO 5 DO
            IF pumpGroup[tmp_i].selection THEN
                pumpGroup[tmp_i].RunComd := TRUE;
            END_IF
        END_FOR
    ELSE
        FOR tmp_i := 1 TO 5 DO
            tmp_priorities[tmp_i] := pumpGroup[tmp_i].priority;
            tmp_pumpIdx[tmp_i] := tmp_i;
        END_FOR
        FOR tmp_i := 1 TO 4 DO
            FOR tmp_j := tmp_i + 1 TO 5 DO
                IF tmp_priorities[tmp_j] > tmp_priorities[tmp_i] THEN
                    tmp_swap := tmp_priorities[tmp_i];
                    tmp_priorities[tmp_i] := tmp_priorities[tmp_j];
                    tmp_priorities[tmp_j] := tmp_swap;
                    tmp_swap_idx := tmp_pumpIdx[tmp_i];
                    tmp_pumpIdx[tmp_i] := tmp_pumpIdx[tmp_j];
                    tmp_pumpIdx[tmp_j] := tmp_swap_idx;
                END_IF
            END_FOR
        END_FOR
        FOR tmp_i := 1 TO 5 DO
            IF tmp_i <= 3 THEN
                pumpGroup[tmp_pumpIdx[tmp_i]].RunComd := TRUE;
            ELSE
                pumpGroup[tmp_pumpIdx[tmp_i]].RunComd := FALSE;
            END_IF
        END_FOR
    END_IF
END_IF

tmp_startPrev := start;
END_FUNCTION_BLOCK

(* ---- public-medium-01.raw_candidate_03.st ---- *)
TYPE ST_Pump :
STRUCT
    priority : INT;
    selection : BOOL;
    RunComd : BOOL;
END_STRUCT
END_TYPE

FUNCTION_BLOCK FB_MultiPumpControl
VAR_INPUT
    mode : BOOL;          // FALSE: Manual mode, TRUE: Automatic mode
    start : BOOL;         // Start button
    stop : BOOL;          // Stop button
END_VAR

VAR_IN_OUT
    pumpGroup : ARRAY[1..5] OF ST_Pump;
END_VAR

VAR
    startRisingEdge : BOOL;               // Rising edge of start
    tmp_startPrev : BOOL;                 // Previous start state
    tmp_i : INT;                          // Loop counter
    tmp_j : INT;                          // Loop counter
    tmp_swap : INT;                       // Swap variable
    tmp_pumpIdx : ARRAY[1..5] OF INT;    // Pump indices for sorting
    tmp_priorities : ARRAY[1..5] OF INT; // Priority copy for sorting
    tmp_swap_idx : INT;                   // Index swap
END_VAR

// ENGINEERING_CONTRACT:
// PUB001 [L91-265]: mode=FALSE → manual; start activates pumps where selection=TRUE
// PUB001 [L91-265]: mode=TRUE → automatic; start activates top-3 by priority (3-in-2-standby)
// PUB002 [L266-350]: stop halts all pumps; no retention on stop (level-triggered)
// PUB003 [L351-463]: Rising edge on start evaluates selection; stop has same-scan priority
// PUB004 [L464-652]: Only RunComd is written; priority/selection are read-only

(* CONTRACT_RULES [] *)

startRisingEdge := start AND NOT tmp_startPrev;

IF stop THEN
    FOR tmp_i := 1 TO 5 DO
        pumpGroup[tmp_i].RunComd := FALSE;
    END_FOR;
ELSIF startRisingEdge THEN
    IF mode = FALSE THEN
        FOR tmp_i := 1 TO 5 DO
            IF pumpGroup[tmp_i].selection THEN
                pumpGroup[tmp_i].RunComd := TRUE;
            END_IF;
        END_FOR;
    ELSE
        FOR tmp_i := 1 TO 5 DO
            tmp_priorities[tmp_i] := pumpGroup[tmp_i].priority;
            tmp_pumpIdx[tmp_i] := tmp_i;
        END_FOR;
        FOR tmp_i := 1 TO 4 DO
            FOR tmp_j := tmp_i + 1 TO 5 DO
                IF tmp_priorities[tmp_j] > tmp_priorities[tmp_i] THEN
                    tmp_swap := tmp_priorities[tmp_i];
                    tmp_priorities[tmp_i] := tmp_priorities[tmp_j];
                    tmp_priorities[tmp_j] := tmp_swap;
                    tmp_swap_idx := tmp_pumpIdx[tmp_i];
                    tmp_pumpIdx[tmp_i] := tmp_pumpIdx[tmp_j];
                    tmp_pumpIdx[tmp_j] := tmp_swap_idx;
                END_IF;
            END_FOR;
        END_FOR;
        FOR tmp_i := 1 TO 5 DO
            IF tmp_i <= 3 THEN
                pumpGroup[tmp_pumpIdx[tmp_i]].RunComd := TRUE;
            ELSE
                pumpGroup[tmp_pumpIdx[tmp_i]].RunComd := FALSE;
            END_IF;
        END_FOR;
    END_IF;
END_IF;

tmp_startPrev := start;
END_FUNCTION_BLOCK

(* ---- public-medium-02.candidate_01.st ---- *)
{attribute 'hide'}
TYPE ST_AnalogChannel : STRUCT
    enable        : BOOL;
    hiLIM         : REAL;
    loLIM         : REAL;
    bipolar       : BOOL;
    measuringMode : INT;
    retVal        : WORD;
    outputValue   : REAL;
END_STRUCT
END_TYPE

FUNCTION_BLOCK FB_AnalogBatchProcessing
VAR_INPUT
END_VAR
VAR_IN_OUT
    count        : DINT;
    analogValues : ARRAY[*] OF INT;
    channels     : ARRAY[*] OF ST_AnalogChannel;
END_VAR
VAR
    tmp_i        : DINT;
    tmp_base     : DINT;
    tmp_raw      : INT;
    tmp_norm     : REAL;
END_VAR

(*
ENGINEERING_CONTRACT
================================================================================
| Output/State      | Activation         | Retention     | Reset          | Scan  | Units           |
|-------------------|--------------------|---------------|----------------|-------|-----------------|
| channels[].retVal | Every enabled chan | Per-call clear| Caller clears  | Final | 16#hex status   |
| channels[].outputValue | Every enabled chan | Caller retains | Caller clears  | Final | REAL engineering|
|-------------------|--------------------|---------------|----------------|-------|-----------------|
PUB001: Process count channels from ordinal position 0 of each array.
PUB002: measuringMode 0=linear(bipolar selectable), 1=stdTemp(raw/10), 2=climTemp(raw/100).
PUB003: Invalid measuringMode -> retVal=16#8001, skip conversion.
PUB004: hiLIM <= loLIM -> retVal=16#8002, skip conversion.
PUB005: Non-temperature linear: unipolar 0..27648->loLIM..hiLIM; bipolar -27648..27648->loLIM..hiLIM.
PUB006: Standard temperature: outputValue = raw * 0.1.
PUB007: Climatic temperature: outputValue = raw * 0.01.
PUB008: Caller provides count 0..min(array lengths); arrays matched by ordinal position.
================================================================================
CONTRACT_RULES []
*)

tmp_base := LOWER_BOUND(analogValues, 1);

FOR tmp_i := 0 TO count - 1 DO
    IF NOT channels[tmp_base + tmp_i].enable THEN
        CONTINUE; // Skip disabled channel
    END_IF

    // Validate measuringMode
    IF channels[tmp_base + tmp_i].measuringMode < 0 OR channels[tmp_base + tmp_i].measuringMode > 2 THEN
        channels[tmp_base + tmp_i].retVal := 16#8001;
        CONTINUE;
    END_IF

    // Validate range
    IF channels[tmp_base + tmp_i].hiLIM <= channels[tmp_base + tmp_i].loLIM THEN
        channels[tmp_base + tmp_i].retVal := 16#8002;
        CONTINUE;
    END_IF

    tmp_raw := analogValues[tmp_base + tmp_i];

    CASE channels[tmp_base + tmp_i].measuringMode OF
        0: // Non-temperature linear scaling
            IF channels[tmp_base + tmp_i].bipolar THEN
                // Bipolar: -27648..27648 -> loLIM..hiLIM
                tmp_norm := INT_TO_REAL(tmp_raw + 27648) / 55296.0;
            ELSE
                // Unipolar: 0..27648 -> loLIM..hiLIM
                tmp_norm := INT_TO_REAL(tmp_raw) / 27648.0;
            END_IF
            channels[tmp_base + tmp_i].outputValue := channels[tmp_base + tmp_i].loLIM + tmp_norm * (channels[tmp_base + tmp_i].hiLIM - channels[tmp_base + tmp_i].loLIM);
            channels[tmp_base + tmp_i].retVal := 16#0000;

        1: // Standard temperature: raw / 10
            channels[tmp_base + tmp_i].outputValue := INT_TO_REAL(tmp_raw) / 10.0;
            channels[tmp_base + tmp_i].retVal := 16#0000;

        2: // Climatic temperature: raw / 100
            channels[tmp_base + tmp_i].outputValue := INT_TO_REAL(tmp_raw) / 100.0;
            channels[tmp_base + tmp_i].retVal := 16#0000;
    END_CASE;
END_FOR;

END_FUNCTION_BLOCK

(* ---- public-medium-02.raw_candidate_01.st ---- *)
{attribute 'hide'}
TYPE ST_AnalogChannel : STRUCT
    enable        : BOOL;
    hiLIM         : REAL;
    loLIM         : REAL;
    bipolar       : BOOL;
    measuringMode : INT;
    retVal        : WORD;
    outputValue   : REAL;
END_STRUCT
END_TYPE

FUNCTION_BLOCK FB_AnalogBatchProcessing
VAR_INPUT
END_VAR
VAR_IN_OUT
    count        : DINT;
    analogValues : ARRAY[*] OF INT;
    channels     : ARRAY[*] OF ST_AnalogChannel;
END_VAR
VAR
    tmp_i        : DINT;
    tmp_base     : DINT;
    tmp_raw      : INT;
    tmp_norm     : REAL;
END_VAR

(*
ENGINEERING_CONTRACT
================================================================================
| Output/State      | Activation         | Retention     | Reset          | Scan  | Units           |
|-------------------|--------------------|---------------|----------------|-------|-----------------|
| channels[].retVal | Every enabled chan | Per-call clear| Caller clears  | Final | 16#hex status   |
| channels[].outputValue | Every enabled chan | Caller retains | Caller clears  | Final | REAL engineering|
|-------------------|--------------------|---------------|----------------|-------|-----------------|
PUB001: Process count channels from ordinal position 0 of each array.
PUB002: measuringMode 0=linear(bipolar selectable), 1=stdTemp(raw/10), 2=climTemp(raw/100).
PUB003: Invalid measuringMode -> retVal=16#8001, skip conversion.
PUB004: hiLIM <= loLIM -> retVal=16#8002, skip conversion.
PUB005: Non-temperature linear: unipolar 0..27648->loLIM..hiLIM; bipolar -27648..27648->loLIM..hiLIM.
PUB006: Standard temperature: outputValue = raw * 0.1.
PUB007: Climatic temperature: outputValue = raw * 0.01.
PUB008: Caller provides count 0..min(array lengths); arrays matched by ordinal position.
================================================================================
CONTRACT_RULES []
*)

tmp_base := LOWER_BOUND(analogValues, 1);

FOR tmp_i := 0 TO count - 1 DO
    IF NOT channels[tmp_base + tmp_i].enable THEN
        CONTINUE; // Skip disabled channel
    END_IF

    // Validate measuringMode
    IF channels[tmp_base + tmp_i].measuringMode < 0 OR channels[tmp_base + tmp_i].measuringMode > 2 THEN
        channels[tmp_base + tmp_i].retVal := 16#8001;
        CONTINUE;
    END_IF

    // Validate range
    IF channels[tmp_base + tmp_i].hiLIM <= channels[tmp_base + tmp_i].loLIM THEN
        channels[tmp_base + tmp_i].retVal := 16#8002;
        CONTINUE;
    END_IF

    tmp_raw := analogValues[tmp_base + tmp_i];

    CASE channels[tmp_base + tmp_i].measuringMode OF
        0: // Non-temperature linear scaling
            IF channels[tmp_base + tmp_i].bipolar THEN
                // Bipolar: -27648..27648 -> loLIM..hiLIM
                tmp_norm := INT_TO_REAL(tmp_raw + 27648) / 55296.0;
            ELSE
                // Unipolar: 0..27648 -> loLIM..hiLIM
                tmp_norm := INT_TO_REAL(tmp_raw) / 27648.0;
            END_IF
            channels[tmp_base + tmp_i].outputValue := channels[tmp_base + tmp_i].loLIM + tmp_norm * (channels[tmp_base + tmp_i].hiLIM - channels[tmp_base + tmp_i].loLIM);
            channels[tmp_base + tmp_i].retVal := 16#0000;

        1: // Standard temperature: raw / 10
            channels[tmp_base + tmp_i].outputValue := INT_TO_REAL(tmp_raw) / 10.0;
            channels[tmp_base + tmp_i].retVal := 16#0000;

        2: // Climatic temperature: raw / 100
            channels[tmp_base + tmp_i].outputValue := INT_TO_REAL(tmp_raw) / 100.0;
            channels[tmp_base + tmp_i].retVal := 16#0000;
    END_CASE;
END_FOR;

END_FUNCTION_BLOCK

(* ---- public-medium-03.candidate_01.st ---- *)
(* ENGINEERING_CONTRACT
+----------------------------------------------------------------+
| Output/State | Activation          | Retention    | Reset       |
+----------------------------------------------------------------+
| average      | New value sampled   | HOLD         | reset=TRUE  |
| windowSizeReached | Window full   | HOLD         | reset=TRUE  |
| error        | windowSize invalid  | LATCHED      | reset=TRUE  |
| status       | Per-error condition | LATCHED      | reset=TRUE  |
+----------------------------------------------------------------+
| Same-scan priority: cyclicExecution > trigger rising edge      |
| Units: windowSize [1..100] slots; average [LREAL]              |
| Boundaries: sampleCount min=0 max=windowSize; index wraps 1-N  |
| Reset priority: reset=TRUE overrides all other inputs          |
| Error condition: windowSize < 1 OR windowSize > 100            |
| Status codes: 16#0000=OK, 16#8200=window size error            |
| Implementation: circular buffer with oldest-value replacement  |
+----------------------------------------------------------------+
*)
(* CONTRACT_RULES [] *)
FUNCTION_BLOCK FB_MovingAverage
VAR_INPUT
    cyclicExecution : BOOL;
    trigger : BOOL;
    value   : LREAL;
    windowSize : INT;
    reset   : BOOL;
END_VAR
VAR_OUTPUT
    average : LREAL;
    windowSizeReached : BOOL;
    error   : BOOL;
    status  : WORD;
END_VAR
VAR
    buffer : ARRAY[1..100] OF LREAL;
    writeIndex : INT := 0;
    sampleCount : INT := 0;
    sum : LREAL := 0.0;
    prevTrigger : BOOL := FALSE;
    tmpValid : BOOL;
    tmpRising : BOOL;
    tmpOldSlot : INT;
END_VAR

tmpValid := (windowSize >= 1) AND (windowSize <= 100);

IF tmpValid THEN
    error := FALSE;
    status := 16#0000;

    IF reset THEN
        writeIndex := 0;
        sampleCount := 0;
        sum := 0.0;
        average := 0.0;
        windowSizeReached := FALSE;
    ELSIF cyclicExecution OR (trigger AND NOT prevTrigger) THEN
        tmpRising := trigger AND NOT prevTrigger;

        IF sampleCount >= windowSize THEN
            tmpOldSlot := ((writeIndex - windowSize) MOD windowSize) + 1;
            sum := sum - buffer[tmpOldSlot];
            sampleCount := sampleCount - 1;
        END_IF;

        writeIndex := (writeIndex MOD windowSize) + 1;
        buffer[writeIndex] := value;
        sum := sum + value;
        sampleCount := sampleCount + 1;

        IF sampleCount > 0 THEN
            average := sum / TO_LREAL(sampleCount);
        END_IF;

        windowSizeReached := (sampleCount >= windowSize);
    END_IF;

    prevTrigger := trigger;
ELSE
    error := TRUE;
    status := 16#8200;
END_IF;

END_FUNCTION_BLOCK

(* ---- public-medium-03.candidate_02.st ---- *)
(* ENGINEERING_CONTRACT
+----------------------------------------------------------------+
| Output/State | Activation          | Retention    | Reset       |
+----------------------------------------------------------------+
| average      | New value sampled   | HOLD         | reset=TRUE  |
| windowSizeReached | Window full   | HOLD         | reset=TRUE  |
| error        | windowSize invalid  | LATCHED      | reset=TRUE  |
| status       | Per-error condition | LATCHED      | reset=TRUE  |
+----------------------------------------------------------------+
| Same-scan priority: cyclicExecution > trigger rising edge      |
| Units: windowSize [1..100] slots; average [LREAL]              |
| Boundaries: sampleCount min=0 max=windowSize; index wraps 1-N  |
| Reset priority: reset=TRUE overrides all other inputs          |
| Error condition: windowSize < 1 OR windowSize > 100            |
| Status codes: 16#0000=OK, 16#8200=window size error            |
| Implementation: circular buffer with oldest-value replacement  |
+----------------------------------------------------------------+
*)
(* CONTRACT_RULES [] *)
FUNCTION_BLOCK FB_MovingAverage
VAR_INPUT
    cyclicExecution : BOOL;
    trigger : BOOL;
    value   : LREAL;
    windowSize : INT;
    reset   : BOOL;
END_VAR
VAR_OUTPUT
    average : LREAL;
    windowSizeReached : BOOL;
    error   : BOOL;
    status  : WORD;
END_VAR
VAR
    buffer : ARRAY[1..100] OF LREAL;
    writeIndex : INT := 0;
    sampleCount : INT := 0;
    sum : LREAL := 0.0;
    prevTrigger : BOOL := FALSE;
    prevWindowSize : INT := 0;
    tmpValid : BOOL;
    tmpRising : BOOL;
    tmpOldSlot : INT;
END_VAR

tmpValid := (windowSize >= 1) AND (windowSize <= 100);

IF tmpValid THEN
    error := FALSE;
    status := 16#0000;

    IF windowSize <> prevWindowSize THEN
        writeIndex := 0;
        sampleCount := 0;
        sum := 0.0;
        windowSizeReached := FALSE;
        prevWindowSize := windowSize;
    END_IF;

    IF reset THEN
        writeIndex := 0;
        sampleCount := 0;
        sum := 0.0;
        average := 0.0;
        windowSizeReached := FALSE;
    ELSIF cyclicExecution OR (trigger AND NOT prevTrigger) THEN
        tmpRising := trigger AND NOT prevTrigger;

        IF sampleCount >= windowSize THEN
            tmpOldSlot := ((writeIndex - windowSize) MOD windowSize) + 1;
            sum := sum - buffer[tmpOldSlot];
            sampleCount := sampleCount - 1;
        END_IF;

        writeIndex := (writeIndex MOD windowSize) + 1;
        buffer[writeIndex] := value;
        sum := sum + value;
        sampleCount := sampleCount + 1;

        IF sampleCount > 0 THEN
            average := sum / TO_LREAL(sampleCount);
        END_IF;

        windowSizeReached := (sampleCount >= windowSize);
    END_IF;

    prevTrigger := trigger;
ELSE
    error := TRUE;
    status := 16#8200;
END_IF;

END_FUNCTION_BLOCK

(* ---- public-medium-03.patch_base_02.st ---- *)
(* ENGINEERING_CONTRACT
+----------------------------------------------------------------+
| Output/State | Activation          | Retention    | Reset       |
+----------------------------------------------------------------+
| average      | New value sampled   | HOLD         | reset=TRUE  |
| windowSizeReached | Window full   | HOLD         | reset=TRUE  |
| error        | windowSize invalid  | LATCHED      | reset=TRUE  |
| status       | Per-error condition | LATCHED      | reset=TRUE  |
+----------------------------------------------------------------+
| Same-scan priority: cyclicExecution > trigger rising edge      |
| Units: windowSize [1..100] slots; average [LREAL]              |
| Boundaries: sampleCount min=0 max=windowSize; index wraps 1-N  |
| Reset priority: reset=TRUE overrides all other inputs          |
| Error condition: windowSize < 1 OR windowSize > 100            |
| Status codes: 16#0000=OK, 16#8200=window size error            |
| Implementation: circular buffer with oldest-value replacement  |
+----------------------------------------------------------------+
*)
(* CONTRACT_RULES [] *)
FUNCTION_BLOCK FB_MovingAverage
VAR_INPUT
    cyclicExecution : BOOL;
    trigger : BOOL;
    value   : LREAL;
    windowSize : INT;
    reset   : BOOL;
END_VAR
VAR_OUTPUT
    average : LREAL;
    windowSizeReached : BOOL;
    error   : BOOL;
    status  : WORD;
END_VAR
VAR
    buffer : ARRAY[1..100] OF LREAL;
    writeIndex : INT := 0;
    sampleCount : INT := 0;
    sum : LREAL := 0.0;
    prevTrigger : BOOL := FALSE;
    tmpValid : BOOL;
    tmpRising : BOOL;
    tmpOldSlot : INT;
END_VAR

tmpValid := (windowSize >= 1) AND (windowSize <= 100);

IF tmpValid THEN
    error := FALSE;
    status := 16#0000;

    IF reset THEN
        writeIndex := 0;
        sampleCount := 0;
        sum := 0.0;
        average := 0.0;
        windowSizeReached := FALSE;
    ELSIF cyclicExecution OR (trigger AND NOT prevTrigger) THEN
        tmpRising := trigger AND NOT prevTrigger;

        IF sampleCount >= windowSize THEN
            tmpOldSlot := ((writeIndex - windowSize) MOD windowSize) + 1;
            sum := sum - buffer[tmpOldSlot];
            sampleCount := sampleCount - 1;
        END_IF;

        writeIndex := (writeIndex MOD windowSize) + 1;
        buffer[writeIndex] := value;
        sum := sum + value;
        sampleCount := sampleCount + 1;

        IF sampleCount > 0 THEN
            average := sum / TO_LREAL(sampleCount);
        END_IF;

        windowSizeReached := (sampleCount >= windowSize);
    END_IF;

    prevTrigger := trigger;
ELSE
    error := TRUE;
    status := 16#8200;
END_IF;

END_FUNCTION_BLOCK

(* ---- public-medium-03.patch_base_03.st ---- *)
(* ENGINEERING_CONTRACT
+----------------------------------------------------------------+
| Output/State | Activation          | Retention    | Reset       |
+----------------------------------------------------------------+
| average      | New value sampled   | HOLD         | reset=TRUE  |
| windowSizeReached | Window full   | HOLD         | reset=TRUE  |
| error        | windowSize invalid  | LATCHED      | reset=TRUE  |
| status       | Per-error condition | LATCHED      | reset=TRUE  |
+----------------------------------------------------------------+
| Same-scan priority: cyclicExecution > trigger rising edge      |
| Units: windowSize [1..100] slots; average [LREAL]              |
| Boundaries: sampleCount min=0 max=windowSize; index wraps 1-N  |
| Reset priority: reset=TRUE overrides all other inputs          |
| Error condition: windowSize < 1 OR windowSize > 100            |
| Status codes: 16#0000=OK, 16#8200=window size error            |
| Implementation: circular buffer with oldest-value replacement  |
+----------------------------------------------------------------+
*)
(* CONTRACT_RULES [] *)
FUNCTION_BLOCK FB_MovingAverage
VAR_INPUT
    cyclicExecution : BOOL;
    trigger : BOOL;
    value   : LREAL;
    windowSize : INT;
    reset   : BOOL;
END_VAR
VAR_OUTPUT
    average : LREAL;
    windowSizeReached : BOOL;
    error   : BOOL;
    status  : WORD;
END_VAR
VAR
    buffer : ARRAY[1..100] OF LREAL;
    writeIndex : INT := 0;
    sampleCount : INT := 0;
    sum : LREAL := 0.0;
    prevTrigger : BOOL := FALSE;
    prevWindowSize : INT := 0;
    tmpValid : BOOL;
    tmpRising : BOOL;
    tmpOldSlot : INT;
END_VAR

tmpValid := (windowSize >= 1) AND (windowSize <= 100);

IF tmpValid THEN
    error := FALSE;
    status := 16#0000;

    IF windowSize <> prevWindowSize THEN
        writeIndex := 0;
        sampleCount := 0;
        sum := 0.0;
        windowSizeReached := FALSE;
        prevWindowSize := windowSize;
    END_IF;

    IF reset THEN
        writeIndex := 0;
        sampleCount := 0;
        sum := 0.0;
        average := 0.0;
        windowSizeReached := FALSE;
    ELSIF cyclicExecution OR (trigger AND NOT prevTrigger) THEN
        tmpRising := trigger AND NOT prevTrigger;

        IF sampleCount >= windowSize THEN
            tmpOldSlot := ((writeIndex - windowSize) MOD windowSize) + 1;
            sum := sum - buffer[tmpOldSlot];
            sampleCount := sampleCount - 1;
        END_IF;

        writeIndex := (writeIndex MOD windowSize) + 1;
        buffer[writeIndex] := value;
        sum := sum + value;
        sampleCount := sampleCount + 1;

        IF sampleCount > 0 THEN
            average := sum / TO_LREAL(sampleCount);
        END_IF;

        windowSizeReached := (sampleCount >= windowSize);
    END_IF;

    prevTrigger := trigger;
ELSE
    error := TRUE;
    status := 16#8200;
END_IF;

END_FUNCTION_BLOCK

(* ---- public-medium-03.patch_base_04.st ---- *)
(* ENGINEERING_CONTRACT
+----------------------------------------------------------------+
| Output/State | Activation          | Retention    | Reset       |
+----------------------------------------------------------------+
| average      | New value sampled   | HOLD         | reset=TRUE  |
| windowSizeReached | Window full   | HOLD         | reset=TRUE  |
| error        | windowSize invalid  | LATCHED      | reset=TRUE  |
| status       | Per-error condition | LATCHED      | reset=TRUE  |
+----------------------------------------------------------------+
| Same-scan priority: cyclicExecution > trigger rising edge      |
| Units: windowSize [1..100] slots; average [LREAL]              |
| Boundaries: sampleCount min=0 max=windowSize; index wraps 1-N  |
| Reset priority: reset=TRUE overrides all other inputs          |
| Error condition: windowSize < 1 OR windowSize > 100            |
| Status codes: 16#0000=OK, 16#8200=window size error            |
| Implementation: circular buffer with oldest-value replacement  |
+----------------------------------------------------------------+
*)
(* CONTRACT_RULES [] *)
FUNCTION_BLOCK FB_MovingAverage
VAR_INPUT
    cyclicExecution : BOOL;
    trigger : BOOL;
    value   : LREAL;
    windowSize : INT;
    reset   : BOOL;
END_VAR
VAR_OUTPUT
    average : LREAL;
    windowSizeReached : BOOL;
    error   : BOOL;
    status  : WORD;
END_VAR
VAR
    buffer : ARRAY[1..100] OF LREAL;
    writeIndex : INT := 0;
    sampleCount : INT := 0;
    sum : LREAL := 0.0;
    prevTrigger : BOOL := FALSE;
    prevWindowSize : INT := 0;
    tmpValid : BOOL;
    tmpRising : BOOL;
    tmpOldSlot : INT;
END_VAR

tmpValid := (windowSize >= 1) AND (windowSize <= 100);

IF tmpValid THEN
    error := FALSE;
    status := 16#0000;

    IF windowSize <> prevWindowSize THEN
        writeIndex := 0;
        sampleCount := 0;
        sum := 0.0;
        windowSizeReached := FALSE;
        prevWindowSize := windowSize;
    END_IF;

    IF reset THEN
        writeIndex := 0;
        sampleCount := 0;
        sum := 0.0;
        average := 0.0;
        windowSizeReached := FALSE;
    ELSIF cyclicExecution OR (trigger AND NOT prevTrigger) THEN
        tmpRising := trigger AND NOT prevTrigger;

        IF sampleCount >= windowSize THEN
            tmpOldSlot := ((writeIndex - windowSize) MOD windowSize) + 1;
            sum := sum - buffer[tmpOldSlot];
            sampleCount := sampleCount - 1;
        END_IF;

        writeIndex := (writeIndex MOD windowSize) + 1;
        buffer[writeIndex] := value;
        sum := sum + value;
        sampleCount := sampleCount + 1;

        IF sampleCount > 0 THEN
            average := sum / TO_LREAL(sampleCount);
        END_IF;

        windowSizeReached := (sampleCount >= windowSize);
    END_IF;

    prevTrigger := trigger;
ELSE
    error := TRUE;
    status := 16#8200;
END_IF;

END_FUNCTION_BLOCK

(* ---- public-medium-03.raw_candidate_01.st ---- *)
(* ENGINEERING_CONTRACT
+----------------------------------------------------------------+
| Output/State | Activation          | Retention    | Reset       |
+----------------------------------------------------------------+
| average      | New value sampled   | HOLD         | reset=TRUE  |
| windowSizeReached | Window full   | HOLD         | reset=TRUE  |
| error        | windowSize invalid  | LATCHED      | reset=TRUE  |
| status       | Per-error condition | LATCHED      | reset=TRUE  |
+----------------------------------------------------------------+
| Same-scan priority: cyclicExecution > trigger rising edge      |
| Units: windowSize [1..100] slots; average [LREAL]              |
| Boundaries: sampleCount min=0 max=windowSize; index wraps 1-N  |
| Reset priority: reset=TRUE overrides all other inputs          |
| Error condition: windowSize < 1 OR windowSize > 100            |
| Status codes: 16#0000=OK, 16#8200=window size error            |
| Implementation: circular buffer with oldest-value replacement  |
+----------------------------------------------------------------+
*)
(* CONTRACT_RULES [] *)
FUNCTION_BLOCK FB_MovingAverage
VAR_INPUT
    cyclicExecution : BOOL;
    trigger : BOOL;
    value   : LREAL;
    windowSize : INT;
    reset   : BOOL;
END_VAR
VAR_OUTPUT
    average : LREAL;
    windowSizeReached : BOOL;
    error   : BOOL;
    status  : WORD;
END_VAR
VAR
    buffer : ARRAY[1..100] OF LREAL;
    writeIndex : INT := 0;
    sampleCount : INT := 0;
    sum : LREAL := 0.0;
    prevTrigger : BOOL := FALSE;
    tmpValid : BOOL;
    tmpRising : BOOL;
    tmpOldSlot : INT;
END_VAR

tmpValid := (windowSize >= 1) AND (windowSize <= 100);

IF tmpValid THEN
    error := FALSE;
    status := 16#0000;

    IF reset THEN
        writeIndex := 0;
        sampleCount := 0;
        sum := 0.0;
        average := 0.0;
        windowSizeReached := FALSE;
    ELSIF cyclicExecution OR (trigger AND NOT prevTrigger) THEN
        tmpRising := trigger AND NOT prevTrigger;

        IF sampleCount >= windowSize THEN
            tmpOldSlot := ((writeIndex - windowSize) MOD windowSize) + 1;
            sum := sum - buffer[tmpOldSlot];
            sampleCount := sampleCount - 1;
        END_IF;

        writeIndex := (writeIndex MOD windowSize) + 1;
        buffer[writeIndex] := value;
        sum := sum + value;
        sampleCount := sampleCount + 1;

        IF sampleCount > 0 THEN
            average := sum / TO_LREAL(sampleCount);
        END_IF;

        windowSizeReached := (sampleCount >= windowSize);
    END_IF;

    prevTrigger := trigger;
ELSE
    error := TRUE;
    status := 16#8200;
END_IF;

END_FUNCTION_BLOCK

(* ---- public-medium-03.raw_candidate_02.st ---- *)
(* ENGINEERING_CONTRACT
+----------------------------------------------------------------+
| Output/State | Activation          | Retention    | Reset       |
+----------------------------------------------------------------+
| average      | New value sampled   | HOLD         | reset=TRUE  |
| windowSizeReached | Window full   | HOLD         | reset=TRUE  |
| error        | windowSize invalid  | LATCHED      | reset=TRUE  |
| status       | Per-error condition | LATCHED      | reset=TRUE  |
+----------------------------------------------------------------+
| Same-scan priority: cyclicExecution > trigger rising edge      |
| Units: windowSize [1..100] slots; average [LREAL]              |
| Boundaries: sampleCount min=0 max=windowSize; index wraps 1-N  |
| Reset priority: reset=TRUE overrides all other inputs          |
| Error condition: windowSize < 1 OR windowSize > 100            |
| Status codes: 16#0000=OK, 16#8200=window size error            |
| Implementation: circular buffer with oldest-value replacement  |
+----------------------------------------------------------------+
*)
(* CONTRACT_RULES [] *)
FUNCTION_BLOCK FB_MovingAverage
VAR_INPUT
    cyclicExecution : BOOL;
    trigger : BOOL;
    value   : LREAL;
    windowSize : INT;
    reset   : BOOL;
END_VAR
VAR_OUTPUT
    average : LREAL;
    windowSizeReached : BOOL;
    error   : BOOL;
    status  : WORD;
END_VAR
VAR
    buffer : ARRAY[1..100] OF LREAL;
    writeIndex : INT := 0;
    sampleCount : INT := 0;
    sum : LREAL := 0.0;
    prevTrigger : BOOL := FALSE;
    prevWindowSize : INT := 0;
    tmpValid : BOOL;
    tmpRising : BOOL;
    tmpOldSlot : INT;
END_VAR

tmpValid := (windowSize >= 1) AND (windowSize <= 100);

IF tmpValid THEN
    error := FALSE;
    status := 16#0000;

    IF windowSize <> prevWindowSize THEN
        writeIndex := 0;
        sampleCount := 0;
        sum := 0.0;
        windowSizeReached := FALSE;
        prevWindowSize := windowSize;
    END_IF;

    IF reset THEN
        writeIndex := 0;
        sampleCount := 0;
        sum := 0.0;
        average := 0.0;
        windowSizeReached := FALSE;
    ELSIF cyclicExecution OR (trigger AND NOT prevTrigger) THEN
        tmpRising := trigger AND NOT prevTrigger;

        IF sampleCount >= windowSize THEN
            tmpOldSlot := ((writeIndex - windowSize) MOD windowSize) + 1;
            sum := sum - buffer[tmpOldSlot];
            sampleCount := sampleCount - 1;
        END_IF;

        writeIndex := (writeIndex MOD windowSize) + 1;
        buffer[writeIndex] := value;
        sum := sum + value;
        sampleCount := sampleCount + 1;

        IF sampleCount > 0 THEN
            average := sum / TO_LREAL(sampleCount);
        END_IF;

        windowSizeReached := (sampleCount >= windowSize);
    END_IF;

    prevTrigger := trigger;
ELSE
    error := TRUE;
    status := 16#8200;
END_IF;

END_FUNCTION_BLOCK

(* ---- public-medium-04.candidate_01.st ---- *)
FUNCTION_BLOCK FB_TemperatureControl
VAR_INPUT
    TemperatureSensorInput : REAL;
    SetTemperature : REAL;
END_VAR

VAR_OUTPUT
    CurrentTemperature : REAL;
    SetTempDisplay : REAL;
    HeaterStatus : BOOL;
    OverheatProtection : BOOL;
    HeaterOutput : BOOL;
END_VAR

VAR
    HeaterRuntimeTimer : TON;
    OverheatCooldownTimer : TON;
    tmp_InOverheatProtection : BOOL;
    tmp_SensorFault : BOOL;
END_VAR

(*
ENGINEERING_CONTRACT
================================================================================
| Output/State        | Activation          | Retention/Reset           | Units/Boundaries     |
|---------------------|---------------------|---------------------------|----------------------|
| CurrentTemperature  | Every scan (copy)   | Unchanged when fault      | REAL, no conversion  |
| SetTempDisplay      | Every scan (copy)   | Always updated            | REAL, no conversion  |
| HeaterStatus        | Every scan (AND)    | False on fault or overheat| BOOL, same-scan      |
| OverheatProtection  | tmp_InOverheatProt  | Hold 3s cooldown then OFF | BOOL, timer-driven   |
| HeaterOutput        | temp < set && !prot | Off on fault, >5s prot,   | BOOL, 5s threshold   |
|                     |                     |   or temp >= set          | > not >= per spec    |
================================================================================
PUB001: temp < set triggers heater on
PUB002: temp > set turns heater off
PUB003: >5s continuous heater runtime triggers overheat protection
PUB004: 3s cooldown before overheat protection can be lifted
PUB005: Sensor fault if input < 0 or > 100
PUB006: Display current temp, set temp, heater status, overheat status
PUB007: Heater must be off during sensor fault
PUB008: Heater off during overheat protection until cooldown completes
================================================================================

CONTRACT_RULES []
*)

// Update display outputs every scan
CurrentTemperature := TemperatureSensorInput;
SetTempDisplay := SetTemperature;

// Detect sensor fault: temperature out of valid range [0, 100]
tmp_SensorFault := (TemperatureSensorInput < 0.0) OR (TemperatureSensorInput > 100.0);

// Determine if heater should be on (based on temperature comparison only)
tmp_HeaterShouldBeOn := (NOT tmp_SensorFault) AND (TemperatureSensorInput < SetTemperature);

// Overheat protection state machine
IF NOT tmp_InOverheatProtection THEN
    // Normal operation: check if overheat protection should trigger
    IF tmp_HeaterShouldBeOn THEN
        // Heater is on, start accumulating runtime
        HeaterRuntimeTimer(IN := TRUE, PT := T#5S);
        IF HeaterRuntimeTimer.Q THEN
            // Heater ran for more than 5 seconds continuously
            tmp_InOverheatProtection := TRUE;
            HeaterRuntimeTimer(IN := FALSE);
        END_IF;
    ELSE
        // Heater is off, reset runtime timer
        HeaterRuntimeTimer(IN := FALSE);
    END_IF;
ELSE
    // In overheat protection state, start 3-second cooldown
    HeaterRuntimeTimer(IN := FALSE);
    OverheatCooldownTimer(IN := TRUE, PT := T#3S);
    IF OverheatCooldownTimer.Q THEN
        // Cooldown complete, clear overheat protection
        tmp_InOverheatProtection := FALSE;
        OverheatCooldownTimer(IN := FALSE);
    END_IF;
END_IF;

// Update overheat protection output
OverheatProtection := tmp_InOverheatProtection;

// Calculate final heater output
// HeaterOutput is true when:
//   - Temperature is below setpoint
//   - Not in sensor fault
//   - Not in overheat protection
HeaterOutput := tmp_HeaterShouldBeOn AND (NOT tmp_InOverheatProtection);

// Heater status follows actual heater output
HeaterStatus := HeaterOutput;

END_FUNCTION_BLOCK

(* ---- public-medium-04.candidate_02.st ---- *)
FUNCTION_BLOCK FB_TemperatureControl
VAR_INPUT
    TemperatureSensorInput : REAL;
    SetTemperature : REAL;
END_VAR

VAR_OUTPUT
    CurrentTemperature : REAL;
    SetTempDisplay : REAL;
    HeaterStatus : BOOL;
    OverheatProtection : BOOL;
    HeaterOutput : BOOL;
END_VAR

VAR
    HeaterRuntimeTimer : TON;
    OverheatCooldownTimer : TON;
    tmp_InOverheatProtection : BOOL;
    tmp_SensorFault : BOOL;
    tmp_HeaterShouldBeOn : BOOL;
END_VAR

(*
ENGINEERING_CONTRACT
================================================================================
| Output/State        | Activation          | Retention/Reset           | Units/Boundaries     |
|---------------------|---------------------|---------------------------|----------------------|
| CurrentTemperature  | Every scan (copy)   | Unchanged when fault      | REAL, no conversion  |
| SetTempDisplay      | Every scan (copy)   | Always updated            | REAL, no conversion  |
| HeaterStatus        | Every scan (AND)    | False on fault or overheat| BOOL, same-scan      |
| OverheatProtection  | tmp_InOverheatProt  | Hold 3s cooldown then OFF | BOOL, timer-driven   |
| HeaterOutput        | temp < set && !prot | Off on fault, >5s prot,   | BOOL, 5s threshold   |
|                     |                     |   or temp >= set          | > not >= per spec    |
================================================================================
PUB001: temp < set triggers heater on
PUB002: temp > set turns heater off
PUB003: >5s continuous heater runtime triggers overheat protection
PUB004: 3s cooldown before overheat protection can be lifted
PUB005: Sensor fault if input < 0 or > 100
PUB006: Display current temp, set temp, heater status, overheat status
PUB007: Heater must be off during sensor fault
PUB008: Heater off during overheat protection until cooldown completes
================================================================================

CONTRACT_RULES []
*)

// Update display outputs every scan
CurrentTemperature := TemperatureSensorInput;
SetTempDisplay := SetTemperature;

// Detect sensor fault: temperature out of valid range [0, 100]
tmp_SensorFault := (TemperatureSensorInput < 0.0) OR (TemperatureSensorInput > 100.0);

// Determine if heater should be on (based on temperature comparison only)
tmp_HeaterShouldBeOn := (NOT tmp_SensorFault) AND (TemperatureSensorInput < SetTemperature);

// Overheat protection state machine
IF NOT tmp_InOverheatProtection THEN
    // Normal operation: check if overheat protection should trigger
    IF tmp_HeaterShouldBeOn THEN
        // Heater is on, start accumulating runtime
        HeaterRuntimeTimer(IN := TRUE, PT := T#5S);
        IF HeaterRuntimeTimer.Q THEN
            // Heater ran for more than 5 seconds continuously
            tmp_InOverheatProtection := TRUE;
            HeaterRuntimeTimer(IN := FALSE);
        END_IF;
    ELSE
        // Heater is off, reset runtime timer
        HeaterRuntimeTimer(IN := FALSE);
    END_IF;
ELSE
    // In overheat protection state, start 3-second cooldown
    HeaterRuntimeTimer(IN := FALSE);
    OverheatCooldownTimer(IN := TRUE, PT := T#3S);
    IF OverheatCooldownTimer.Q THEN
        // Cooldown complete, clear overheat protection
        tmp_InOverheatProtection := FALSE;
        OverheatCooldownTimer(IN := FALSE);
    END_IF;
END_IF;

// Update overheat protection output
OverheatProtection := tmp_InOverheatProtection;

// Calculate final heater output
// HeaterOutput is true when:
//   - Temperature is below setpoint
//   - Not in sensor fault
//   - Not in overheat protection
HeaterOutput := tmp_HeaterShouldBeOn AND (NOT tmp_InOverheatProtection);

// Heater status follows actual heater output
HeaterStatus := HeaterOutput;

END_FUNCTION_BLOCK

(* ---- public-medium-04.candidate_04.st ---- *)
FUNCTION_BLOCK FB_TemperatureControl
VAR_INPUT
    TemperatureSensorInput : REAL;
    SetTemperature : REAL;
END_VAR

VAR_OUTPUT
    CurrentTemperature : REAL;
    SetTempDisplay : REAL;
    HeaterStatus : BOOL;
    OverheatProtection : BOOL;
    HeaterOutput : BOOL;
END_VAR

VAR
    HeaterRuntimeTimer : TON;
    OverheatCooldownTimer : TON;
    tmp_InOverheatProtection : BOOL;
    tmp_SensorFault : BOOL;
    tmp_RuntimeTimerEnable : BOOL;
END_VAR

(*
ENGINEERING_CONTRACT
================================================================================
| Output/State        | Activation          | Retention/Reset           | Units/Boundaries     |
|---------------------|---------------------|---------------------------|----------------------|
| CurrentTemperature  | Every scan (copy)   | Unchanged when fault      | REAL, no conversion  |
| SetTempDisplay      | Every scan (copy)   | Always updated            | REAL, no conversion  |
| HeaterStatus        | Every scan (AND)    | False on fault or overheat| BOOL, same-scan      |
| OverheatProtection  | tmp_InOverheatProt  | Hold 3s cooldown then OFF | BOOL, timer-driven   |
| HeaterOutput        | temp < set && !prot | Off on fault, >5s prot,   | BOOL, 5s threshold   |
|                     |                     |   or temp >= set          | > not >= per spec    |
================================================================================
PUB001: temp < set triggers heater on
PUB002: temp > set turns heater off
PUB003: >5s continuous heater runtime triggers overheat protection
PUB004: 3s cooldown before overheat protection can be lifted
PUB005: Sensor fault if input < 0 or > 100
PUB006: Display current temp, set temp, heater status, overheat status
PUB007: Heater must be off during sensor fault
PUB008: Heater off during overheat protection until cooldown completes
================================================================================

CONTRACT_RULES []
*)

// Update display outputs every scan
CurrentTemperature := TemperatureSensorInput;
SetTempDisplay := SetTemperature;

// Detect sensor fault: temperature out of valid range [0, 100]
tmp_SensorFault := (TemperatureSensorInput < 0.0) OR (TemperatureSensorInput > 100.0);

// Determine if runtime timer should accumulate (heater on, not in fault, not in overheat protection)
tmp_RuntimeTimerEnable := (NOT tmp_SensorFault) AND (NOT tmp_InOverheatProtection) AND (TemperatureSensorInput < SetTemperature);

// Overheat protection state machine
IF NOT tmp_InOverheatProtection THEN
    // Normal operation: check if overheat protection should trigger
    IF tmp_RuntimeTimerEnable THEN
        // Heater is on, start accumulating runtime
        HeaterRuntimeTimer(IN := TRUE, PT := T#5001MS);
        IF HeaterRuntimeTimer.Q THEN
            // Heater ran for more than 5 seconds continuously
            tmp_InOverheatProtection := TRUE;
            HeaterRuntimeTimer(IN := FALSE);
        END_IF;
    ELSE
        // Heater is off or in fault, reset runtime timer
        HeaterRuntimeTimer(IN := FALSE);
    END_IF;
ELSE
    // In overheat protection state, run 3-second cooldown
    HeaterRuntimeTimer(IN := FALSE);
    OverheatCooldownTimer(IN := TRUE, PT := T#3S);
    IF OverheatCooldownTimer.Q THEN
        // Cooldown complete, clear overheat protection
        tmp_InOverheatProtection := FALSE;
        OverheatCooldownTimer(IN := FALSE);
    END_IF;
END_IF;

// Update outputs
OverheatProtection := tmp_InOverheatProtection;

// Calculate final heater output: on when temperature below setpoint, not in fault, not in overheat protection
HeaterOutput := tmp_RuntimeTimerEnable;

// Heater status follows actual heater output
HeaterStatus := HeaterOutput;

END_FUNCTION_BLOCK

(* ---- public-medium-04.patch_base_02.st ---- *)
FUNCTION_BLOCK FB_TemperatureControl
VAR_INPUT
    TemperatureSensorInput : REAL;
    SetTemperature : REAL;
END_VAR

VAR_OUTPUT
    CurrentTemperature : REAL;
    SetTempDisplay : REAL;
    HeaterStatus : BOOL;
    OverheatProtection : BOOL;
    HeaterOutput : BOOL;
END_VAR

VAR
    HeaterRuntimeTimer : TON;
    OverheatCooldownTimer : TON;
    tmp_InOverheatProtection : BOOL;
    tmp_SensorFault : BOOL;
END_VAR

(*
ENGINEERING_CONTRACT
================================================================================
| Output/State        | Activation          | Retention/Reset           | Units/Boundaries     |
|---------------------|---------------------|---------------------------|----------------------|
| CurrentTemperature  | Every scan (copy)   | Unchanged when fault      | REAL, no conversion  |
| SetTempDisplay      | Every scan (copy)   | Always updated            | REAL, no conversion  |
| HeaterStatus        | Every scan (AND)    | False on fault or overheat| BOOL, same-scan      |
| OverheatProtection  | tmp_InOverheatProt  | Hold 3s cooldown then OFF | BOOL, timer-driven   |
| HeaterOutput        | temp < set && !prot | Off on fault, >5s prot,   | BOOL, 5s threshold   |
|                     |                     |   or temp >= set          | > not >= per spec    |
================================================================================
PUB001: temp < set triggers heater on
PUB002: temp > set turns heater off
PUB003: >5s continuous heater runtime triggers overheat protection
PUB004: 3s cooldown before overheat protection can be lifted
PUB005: Sensor fault if input < 0 or > 100
PUB006: Display current temp, set temp, heater status, overheat status
PUB007: Heater must be off during sensor fault
PUB008: Heater off during overheat protection until cooldown completes
================================================================================

CONTRACT_RULES []
*)

// Update display outputs every scan
CurrentTemperature := TemperatureSensorInput;
SetTempDisplay := SetTemperature;

// Detect sensor fault: temperature out of valid range [0, 100]
tmp_SensorFault := (TemperatureSensorInput < 0.0) OR (TemperatureSensorInput > 100.0);

// Determine if heater should be on (based on temperature comparison only)
tmp_HeaterShouldBeOn := (NOT tmp_SensorFault) AND (TemperatureSensorInput < SetTemperature);

// Overheat protection state machine
IF NOT tmp_InOverheatProtection THEN
    // Normal operation: check if overheat protection should trigger
    IF tmp_HeaterShouldBeOn THEN
        // Heater is on, start accumulating runtime
        HeaterRuntimeTimer(IN := TRUE, PT := T#5S);
        IF HeaterRuntimeTimer.Q THEN
            // Heater ran for more than 5 seconds continuously
            tmp_InOverheatProtection := TRUE;
            HeaterRuntimeTimer(IN := FALSE);
        END_IF;
    ELSE
        // Heater is off, reset runtime timer
        HeaterRuntimeTimer(IN := FALSE);
    END_IF;
ELSE
    // In overheat protection state, start 3-second cooldown
    HeaterRuntimeTimer(IN := FALSE);
    OverheatCooldownTimer(IN := TRUE, PT := T#3S);
    IF OverheatCooldownTimer.Q THEN
        // Cooldown complete, clear overheat protection
        tmp_InOverheatProtection := FALSE;
        OverheatCooldownTimer(IN := FALSE);
    END_IF;
END_IF;

// Update overheat protection output
OverheatProtection := tmp_InOverheatProtection;

// Calculate final heater output
// HeaterOutput is true when:
//   - Temperature is below setpoint
//   - Not in sensor fault
//   - Not in overheat protection
HeaterOutput := tmp_HeaterShouldBeOn AND (NOT tmp_InOverheatProtection);

// Heater status follows actual heater output
HeaterStatus := HeaterOutput;

END_FUNCTION_BLOCK

(* ---- public-medium-04.patch_base_03.st ---- *)
FUNCTION_BLOCK FB_TemperatureControl
VAR_INPUT
    TemperatureSensorInput : REAL;
    SetTemperature : REAL;
END_VAR

VAR_OUTPUT
    CurrentTemperature : REAL;
    SetTempDisplay : REAL;
    HeaterStatus : BOOL;
    OverheatProtection : BOOL;
    HeaterOutput : BOOL;
END_VAR

VAR
    HeaterRuntimeTimer : TON;
    OverheatCooldownTimer : TON;
    tmp_InOverheatProtection : BOOL;
    tmp_SensorFault : BOOL;
    tmp_HeaterShouldBeOn : BOOL;
END_VAR

(*
ENGINEERING_CONTRACT
================================================================================
| Output/State        | Activation          | Retention/Reset           | Units/Boundaries     |
|---------------------|---------------------|---------------------------|----------------------|
| CurrentTemperature  | Every scan (copy)   | Unchanged when fault      | REAL, no conversion  |
| SetTempDisplay      | Every scan (copy)   | Always updated            | REAL, no conversion  |
| HeaterStatus        | Every scan (AND)    | False on fault or overheat| BOOL, same-scan      |
| OverheatProtection  | tmp_InOverheatProt  | Hold 3s cooldown then OFF | BOOL, timer-driven   |
| HeaterOutput        | temp < set && !prot | Off on fault, >5s prot,   | BOOL, 5s threshold   |
|                     |                     |   or temp >= set          | > not >= per spec    |
================================================================================
PUB001: temp < set triggers heater on
PUB002: temp > set turns heater off
PUB003: >5s continuous heater runtime triggers overheat protection
PUB004: 3s cooldown before overheat protection can be lifted
PUB005: Sensor fault if input < 0 or > 100
PUB006: Display current temp, set temp, heater status, overheat status
PUB007: Heater must be off during sensor fault
PUB008: Heater off during overheat protection until cooldown completes
================================================================================

CONTRACT_RULES []
*)

// Update display outputs every scan
CurrentTemperature := TemperatureSensorInput;
SetTempDisplay := SetTemperature;

// Detect sensor fault: temperature out of valid range [0, 100]
tmp_SensorFault := (TemperatureSensorInput < 0.0) OR (TemperatureSensorInput > 100.0);

// Determine if heater should be on (based on temperature comparison only)
tmp_HeaterShouldBeOn := (NOT tmp_SensorFault) AND (TemperatureSensorInput < SetTemperature);

// Overheat protection state machine
IF NOT tmp_InOverheatProtection THEN
    // Normal operation: check if overheat protection should trigger
    IF tmp_HeaterShouldBeOn THEN
        // Heater is on, start accumulating runtime
        HeaterRuntimeTimer(IN := TRUE, PT := T#5S);
        IF HeaterRuntimeTimer.Q THEN
            // Heater ran for more than 5 seconds continuously
            tmp_InOverheatProtection := TRUE;
            HeaterRuntimeTimer(IN := FALSE);
        END_IF;
    ELSE
        // Heater is off, reset runtime timer
        HeaterRuntimeTimer(IN := FALSE);
    END_IF;
ELSE
    // In overheat protection state, start 3-second cooldown
    HeaterRuntimeTimer(IN := FALSE);
    OverheatCooldownTimer(IN := TRUE, PT := T#3S);
    IF OverheatCooldownTimer.Q THEN
        // Cooldown complete, clear overheat protection
        tmp_InOverheatProtection := FALSE;
        OverheatCooldownTimer(IN := FALSE);
    END_IF;
END_IF;

// Update overheat protection output
OverheatProtection := tmp_InOverheatProtection;

// Calculate final heater output
// HeaterOutput is true when:
//   - Temperature is below setpoint
//   - Not in sensor fault
//   - Not in overheat protection
HeaterOutput := tmp_HeaterShouldBeOn AND (NOT tmp_InOverheatProtection);

// Heater status follows actual heater output
HeaterStatus := HeaterOutput;

END_FUNCTION_BLOCK
